// TwinCAT 3 PLC project MBIDivB_Tests
// ProgramVersion: 3.1.4024.0
// libraries:
//   MBIDivB, * (MBI Div-B)
//   Tc2_Standard, * (Beckhoff Automation GmbH)
//   Tc2_System, * (Beckhoff Automation GmbH)
//   Tc3_Module, * (Beckhoff Automation GmbH)
//   TcUnit, * (www.tcunit.org)
// project tree:
//   Example/ PRG_EXAMPLE.TcPOU
//   POUs/ FB_PlcShutdownTestable.TcPOU, PRG_TEST.TcPOU
//   / PlcTask.TcTTO
//   Tests/ FB_AnalogInputTest.TcPOU, FB_AnalogOutputTest.TcPOU, FB_CounterTimerTest.TcPOU, FB_EndPositionSwitchesTest.TcPOU, FB_FemtoAmplifierTest.TcPOU, FB_FlowMeterTest.TcPOU, FB_LedControlTest.TcPOU, FB_MultiTriggerTest.TcPOU, FB_ParameterTest.TcPOU, FB_PlcShutdownTest.TcPOU, FB_ShutterControlTest.TcPOU, FB_TimeTest.TcPOU
// (motion and I/O tree: see PLC project mbidivb)
// real-time tasks:
//   TASK PlcTask: cycle T#10ms, priority 20, ADS port 350
//   TASK PlcTask1: cycle T#1ms, priority 21, ADS port 351
// variable links:
//   MBIDivB_Tests/MBIDivB_Tests Instance <-> Device 1 (EtherCAT)/Term 1 (EK1100)/EL3102 (EL3102)
//     PlcTask Inputs/PRG_EXAMPLE.Ai1.Raw <-> AI Standard Channel 1/Value
//   MBIDivB_Tests/MBIDivB_Tests Instance <-> Device 1 (EtherCAT)/Term 1 (EK1100)/ELM3142 (ELM3142-0000)
//     PlcTask Inputs/PRG_EXAMPLE.Ai2.Raw <-> PAI Samples 1 Channel 1/Samples[0]
//   MBIDivB_Tests/MBIDivB_Tests Instance <-> Device 1 (EtherCAT)/Term 1 (EK1100)/Term 4 (EL2595)
//     PlcTask Inputs/PRG_EXAMPLE.Led1.InfoData1 <-> DOX Synchron info data/Info data 1
//     PlcTask Inputs/PRG_EXAMPLE.Led1.InfoData2 <-> DOX Synchron info data/Info data 2
//     PlcTask Inputs/PRG_EXAMPLE.Led1.StatusWord <-> DOX Status/Status
//     PlcTask Outputs/PRG_EXAMPLE.Led1.ControlWord <-> DOX Control/Control
//   MBIDivB_Tests/MBIDivB_Tests Instance <-> Device 1 (EtherCAT)/Term 1 (EK1100)/Term 5 (EL2124)
//     PlcTask Outputs/PRG_EXAMPLE.Femto1.GainBit0 <-> Channel 1/Output
//     PlcTask Outputs/PRG_EXAMPLE.Femto1.GainBit1 <-> Channel 2/Output
//     PlcTask Outputs/PRG_EXAMPLE.Femto1.GainBit2 <-> Channel 3/Output
//     PlcTask Outputs/PRG_EXAMPLE.Femto1.LowNoise <-> Channel 4/Output
//   MBIDivB_Tests/MBIDivB_Tests Instance <-> Device 1 (EtherCAT)/Term 1 (EK1100)/Term 6 (EL2124)
//     PlcTask Outputs/PRG_EXAMPLE.Femto1.DcCoupling <-> Channel 1/Output
//   MBIDivB_Tests/MBIDivB_Tests Instance <-> Device 1 (EtherCAT)/Term 1 (EK1100)/Term 7 (EL1124)
//     PlcTask Inputs/PRG_EXAMPLE.Femto1.Overload <-> Channel 1/Input

CONFIGURATION MBIDivB_Tests
    RESOURCE PLC ON TwinCAT3
        TASK PlcTask(INTERVAL := T#1ms, PRIORITY := 21);
        PROGRAM PRG_TEST WITH PlcTask : PRG_TEST;
        PROGRAM PRG_EXAMPLE WITH PlcTask : PRG_EXAMPLE;
    END_RESOURCE
END_CONFIGURATION

// ---- POUs/PRG_TEST.TcPOU

(*
    Runs all MBIDivB test suites with TcUnit. Call it from the test task
    (1 ms cycle time).
*)
PROGRAM PRG_TEST
VAR
    TimeTest : FB_TimeTest;
    ParameterTest : FB_ParameterTest;
    AnalogInputTest : FB_AnalogInputTest;
    CounterTimerTest : FB_CounterTimerTest;
    AnalogOutputTest : FB_AnalogOutputTest;
    MultiTriggerTest : FB_MultiTriggerTest;
    FlowMeterTest : FB_FlowMeterTest;
    ShutterControlTest : FB_ShutterControlTest;
    LedControlTest : FB_LedControlTest;
    FemtoAmplifierTest : FB_FemtoAmplifierTest;
    EndPositionSwitchesTest : FB_EndPositionSwitchesTest;
    PlcShutdownTest : FB_PlcShutdownTest;
END_VAR


TcUnit.RUN();

END_PROGRAM

// ---- Tests/FB_TimeTest.TcPOU

(*
    Tests of F_MsToCyclesAt, F_CyclesToMsAt and the test task's cycle time.
*)
FUNCTION_BLOCK FB_TimeTest EXTENDS TcUnit.FB_TestSuite


TaskCycleTimeIs1ms();
Converts2_4msAt1ms();
Converts1msAt0_3ms();
Converts100msAt10ms();
NonPositiveTimeGivesZero();


METHOD PRIVATE Converts100msAt10ms

TEST('Converts100msAt10ms');

AssertEquals_UDINT(Expected := 10, Actual := MBIDivB.F_MsToCyclesAt(TimeMs := 100.0, CycleTime := 100000), Message := 'cycles');
AssertEquals_REAL(Expected := 100.0, Actual := MBIDivB.F_CyclesToMsAt(Cycles := 10, CycleTime := 100000), Delta := 1.0E-6, Message := 'effective ms');

TEST_FINISHED();
END_METHOD


METHOD PRIVATE Converts1msAt0_3ms

TEST('Converts1msAt0_3ms');

AssertEquals_UDINT(Expected := 3, Actual := MBIDivB.F_MsToCyclesAt(TimeMs := 1.0, CycleTime := 3000), Message := 'cycles');
AssertEquals_REAL(Expected := 0.9, Actual := MBIDivB.F_CyclesToMsAt(Cycles := 3, CycleTime := 3000), Delta := 1.0E-6, Message := 'effective ms');

TEST_FINISHED();
END_METHOD


METHOD PRIVATE Converts2_4msAt1ms

TEST('Converts2_4msAt1ms');

AssertEquals_UDINT(Expected := 2, Actual := MBIDivB.F_MsToCyclesAt(TimeMs := 2.4, CycleTime := 10000), Message := 'cycles');
AssertEquals_REAL(Expected := 2.0, Actual := MBIDivB.F_CyclesToMsAt(Cycles := 2, CycleTime := 10000), Delta := 1.0E-6, Message := 'effective ms');

TEST_FINISHED();
END_METHOD


METHOD PRIVATE NonPositiveTimeGivesZero

TEST('NonPositiveTimeGivesZero');

AssertEquals_UDINT(Expected := 0, Actual := MBIDivB.F_MsToCyclesAt(TimeMs := 0.0, CycleTime := 10000), Message := 'zero');
AssertEquals_UDINT(Expected := 0, Actual := MBIDivB.F_MsToCyclesAt(TimeMs := -5.0, CycleTime := 10000), Message := 'negative');
AssertEquals_UDINT(Expected := 0, Actual := MBIDivB.F_MsToCyclesAt(TimeMs := 5.0, CycleTime := 0), Message := 'cycle time 0');

TEST_FINISHED();
END_METHOD


METHOD PRIVATE TaskCycleTimeIs1ms

TEST('TaskCycleTimeIs1ms');

AssertEquals_UDINT(Expected := 10000, Actual := MBIDivB.F_GetTaskCycleTime(),
    Message := 'The test task must run at 1 ms; the other suites assume it');

TEST_FINISHED();
END_METHOD

END_FUNCTION_BLOCK

// ---- Tests/FB_ParameterTest.TcPOU

(*
    Checks that the library parameter overrides of this test project take
    effect (task 10.1). Expected overrides in the Library Manager:
    CT_CHANNELS 4, CT_BUFFER_LENGTH 1000, AO_WAVEFORM_LENGTH 1000,
    FLOW_BUFFER_LENGTH 100.
*)
FUNCTION_BLOCK FB_ParameterTest EXTENDS TcUnit.FB_TestSuite
VAR
    Ct : MBIDivB.FB_CounterTimer;
    Ao : MBIDivB.FB_AnalogOutput;
END_VAR


OverridesSetArrayBounds();


METHOD PRIVATE OverridesSetArrayBounds

TEST('OverridesSetArrayBounds');

// Element counts from the array sizes (UPPER_BOUND only works on
// variable-length arrays in TwinCAT 3.1.4024).
AssertEquals_UDINT(Expected := 4, Actual := TO_UDINT(SIZEOF(Ct.Channel) / SIZEOF(Ct.Channel[1])), Message := 'CT_CHANNELS');
AssertEquals_UDINT(Expected := 1000, Actual := TO_UDINT(SIZEOF(Ct.Channel[1].Data) / SIZEOF(Ct.Channel[1].Data[1])), Message := 'CT_BUFFER_LENGTH');
AssertEquals_UDINT(Expected := 1000, Actual := TO_UDINT(SIZEOF(Ao.Data) / SIZEOF(Ao.Data[1])), Message := 'AO_WAVEFORM_LENGTH');
AssertEquals_UDINT(Expected := 100, Actual := MBIDivB.GVL_Param.FLOW_BUFFER_LENGTH, Message := 'FLOW_BUFFER_LENGTH');

TEST_FINISHED();
END_METHOD

END_FUNCTION_BLOCK

// ---- Tests/FB_AnalogInputTest.TcPOU

(*
    Tests of FB_AnalogInput16/32 (specs/analog-input).
*)
FUNCTION_BLOCK FB_AnalogInputTest EXTENDS TcUnit.FB_TestSuite
VAR
    AiNegative : MBIDivB.FB_AnalogInput16;
    AiElmNominal : MBIDivB.FB_AnalogInput32;
    AiElmPreset : MBIDivB.FB_AnalogInput32;
    AiZeroScale : MBIDivB.FB_AnalogInput16;
    AiConstant : MBIDivB.FB_AnalogInput16;
    AiReduced : MBIDivB.FB_AnalogInput16;
    AiSizeZero : MBIDivB.FB_AnalogInput16;
    AiOverrange : MBIDivB.FB_AnalogInput16;
    AiUnlinked : MBIDivB.FB_AnalogInput32;
    AiRestartStep : MBIDivB.FB_AnalogInput16;
    AiRestartSettings : MBIDivB.FB_AnalogInput32;
END_VAR


NegativeValue16Bit();
ElmNominalFullScale();
ElmExtendedPreset();
ZeroRawFullScaleRejected();
ConstantInputFiltered();
FilterSizeReducedRestarts();
FilterSizeZeroClampedToOne();
OverrangeSetAndCleared();
UnlinkedStatusBitsNoError();
RestartAfterStep();
RestartKeepsSettings();


METHOD PRIVATE ConstantInputFiltered
VAR
    Cycle : INT;
END_VAR

TEST('ConstantInputFiltered');

AiConstant.SetScale(RawFullScale := 1, ValueFullScale := 1.0);
AiConstant.Cfg.FilterSize := 10;
AiConstant.Raw := 2;
FOR Cycle := 1 TO 25 DO
    AiConstant();
END_FOR
AssertEquals_REAL(Expected := 2.0, Actual := AiConstant.Status.ValueFiltered, Delta := 1.0E-6, Message := 'ValueFiltered');

TEST_FINISHED();
END_METHOD


METHOD PRIVATE ElmExtendedPreset

TEST('ElmExtendedPreset');

AiElmPreset.SetScalePreset(Preset := MBIDivB.E_AiScalePreset.ELM3XXX_EXTENDED, NominalFullScale := 10.0);
AiElmPreset.Raw := 7812500;
AiElmPreset();
AssertEquals_REAL(Expected := 10.0, Actual := AiElmPreset.Status.Value, Delta := 1.0E-5, Message := 'nominal');
AiElmPreset.Raw := 8388607;
AiElmPreset();
AssertEquals_REAL(Expected := 10.737, Actual := AiElmPreset.Status.Value, Delta := 0.001, Message := 'technical full scale');

TEST_FINISHED();
END_METHOD


METHOD PRIVATE ElmNominalFullScale

TEST('ElmNominalFullScale');

AiElmNominal.SetScale(RawFullScale := 7812500, ValueFullScale := 10.0);
AiElmNominal.Raw := 7812500;
AiElmNominal();
AssertEquals_REAL(Expected := 10.0, Actual := AiElmNominal.Status.Value, Delta := 1.0E-5, Message := 'Value');
AssertEquals_DINT(Expected := 7812500, Actual := AiElmNominal.Status.RawFullScale, Message := 'RawFullScale');
AssertEquals_REAL(Expected := 10.0, Actual := AiElmNominal.Status.ValueFullScale, Delta := 1.0E-6, Message := 'ValueFullScale');

TEST_FINISHED();
END_METHOD


METHOD PRIVATE FilterSizeReducedRestarts
VAR
    Cycle : INT;
END_VAR

TEST('FilterSizeReducedRestarts');

AiReduced.SetScale(RawFullScale := 1, ValueFullScale := 1.0);
AiReduced.Cfg.FilterSize := 1000;
AiReduced.Raw := 3;
FOR Cycle := 1 TO 100 DO
    AiReduced();
END_FOR
AiReduced.Cfg.FilterSize := 10;
AiReduced.Raw := 1;
AiReduced();
AssertEquals_REAL(Expected := 1.0, Actual := AiReduced.Status.ValueFiltered, Delta := 1.0E-6, Message := 'no contribution from older samples');

TEST_FINISHED();
END_METHOD


METHOD PRIVATE FilterSizeZeroClampedToOne

TEST('FilterSizeZeroClampedToOne');

AiSizeZero.SetScale(RawFullScale := 1, ValueFullScale := 1.0);
AiSizeZero.Cfg.FilterSize := 0;
AiSizeZero.Raw := 4;
AiSizeZero();
AssertEquals_DINT(Expected := 1, Actual := AiSizeZero.Cfg.FilterSize, Message := 'FilterSize written back');
AssertEquals_REAL(Expected := 4.0, Actual := AiSizeZero.Status.ValueFiltered, Delta := 1.0E-6, Message := 'ValueFiltered');

TEST_FINISHED();
END_METHOD


METHOD PRIVATE NegativeValue16Bit

TEST('NegativeValue16Bit');

AiNegative.SetScalePreset(Preset := MBIDivB.E_AiScalePreset.EL31XX_LEGACY, NominalFullScale := 10.0);
AiNegative.Raw := -16384;
AiNegative();
AssertEquals_REAL(Expected := -5.0, Actual := AiNegative.Status.Value, Delta := 0.001, Message := 'Value');
AssertEquals_DINT(Expected := -16384, Actual := AiNegative.Status.Raw, Message := 'Raw');

TEST_FINISHED();
END_METHOD


METHOD PRIVATE OverrangeSetAndCleared

TEST('OverrangeSetAndCleared');

AiOverrange.Overrange := TRUE;
AiOverrange();
AssertTrue(Condition := AiOverrange.Status.Error, Message := 'Error while set');
AssertTrue(Condition := FIND(AiOverrange.Status.ErrorText, 'overrange') > 0, Message := 'ErrorText mentions overrange');
AiOverrange.Overrange := FALSE;
AiOverrange();
AssertFalse(Condition := AiOverrange.Status.Error, Message := 'Error cleared');
AssertEquals_STRING(Expected := '', Actual := AiOverrange.Status.ErrorText, Message := 'ErrorText cleared');

TEST_FINISHED();
END_METHOD


METHOD PRIVATE RestartAfterStep
VAR
    Cycle : INT;
    Wrong : INT;
END_VAR

TEST('RestartAfterStep');

AiRestartStep.SetScale(RawFullScale := 1000, ValueFullScale := 1.0);
AiRestartStep.Cfg.FilterSize := 10;
AiRestartStep.Raw := 1000;
FOR Cycle := 1 TO 15 DO
    AiRestartStep();
END_FOR
AiRestartStep.RestartFilter();
AiRestartStep.Raw := 3000;
FOR Cycle := 1 TO 12 DO
    AiRestartStep();
    IF ABS(AiRestartStep.Status.ValueFiltered - 3.0) > 1.0E-6 THEN
        Wrong := Wrong + 1;
    END_IF
END_FOR
AssertEquals_INT(Expected := 0, Actual := Wrong, Message := 'calls with ValueFiltered <> 3.0 V after the restart');

TEST_FINISHED();
END_METHOD


METHOD PRIVATE RestartKeepsSettings

TEST('RestartKeepsSettings');

AiRestartSettings.SetScale(RawFullScale := 7812500, ValueFullScale := 10.0);
AiRestartSettings.Cfg.FilterSize := 20;
AiRestartSettings.Raw := 3906250;
AiRestartSettings();
AiRestartSettings.RestartFilter();
AiRestartSettings();
AssertEquals_DINT(Expected := 20, Actual := AiRestartSettings.Cfg.FilterSize, Message := 'FilterSize');
AssertEquals_DINT(Expected := 7812500, Actual := AiRestartSettings.Status.RawFullScale, Message := 'RawFullScale');
AssertEquals_REAL(Expected := 10.0, Actual := AiRestartSettings.Status.ValueFullScale, Delta := 1.0E-6, Message := 'ValueFullScale');
AssertEquals_REAL(Expected := 5.0, Actual := AiRestartSettings.Status.Value, Delta := 1.0E-5, Message := 'Value');

TEST_FINISHED();
END_METHOD


METHOD PRIVATE UnlinkedStatusBitsNoError

TEST('UnlinkedStatusBitsNoError');

AiUnlinked.Raw := 1000;
AiUnlinked();
AssertFalse(Condition := AiUnlinked.Status.Error, Message := 'Error');

TEST_FINISHED();
END_METHOD


METHOD PRIVATE ZeroRawFullScaleRejected
VAR
    Accepted : BOOL;
END_VAR

TEST('ZeroRawFullScaleRejected');

AiZeroScale.SetScale(RawFullScale := 32767, ValueFullScale := 10.0);
Accepted := AiZeroScale.SetScale(RawFullScale := 0, ValueFullScale := 5.0);
AiZeroScale.Raw := 16384;
AiZeroScale();
AssertFalse(Condition := Accepted, Message := 'SetScale must return FALSE');
AssertTrue(Condition := AiZeroScale.Status.Error, Message := 'Error');
AssertTrue(Condition := FIND(AiZeroScale.Status.ErrorText, 'RawFullScale') > 0, Message := 'ErrorText names RawFullScale');
AssertEquals_REAL(Expected := 5.0, Actual := AiZeroScale.Status.Value, Delta := 0.001, Message := 'previous scaling kept');

TEST_FINISHED();
END_METHOD

END_FUNCTION_BLOCK

// ---- Tests/FB_CounterTimerTest.TcPOU

(*
    Tests of FB_CounterTimer (specs/counter-timer) and of the command
    handshake and error rules (specs/ads-interface) on this block.
    Needs CT_CHANNELS >= 4.
*)
FUNCTION_BLOCK FB_CounterTimerTest EXTENDS TcUnit.FB_TestSuite
VAR
    CtSync : MBIDivB.FB_CounterTimer;
    CtTooMany : MBIDivB.FB_CounterTimer;
    CtLinear : MBIDivB.FB_CounterTimer;
    CtLatency : MBIDivB.FB_CounterTimer;
    CtTrigger : MBIDivB.FB_CounterTimer;
    CtMissed : MBIDivB.FB_CounterTimer;
    CtProgress : MBIDivB.FB_CounterTimer;
    CtStop : MBIDivB.FB_CounterTimer;
    CtRunning : MBIDivB.FB_CounterTimer;
    CtHandshake : MBIDivB.FB_CounterTimer;
    CtErrorClear : MBIDivB.FB_CounterTimer;
    CtCfgChange : MBIDivB.FB_CounterTimer;
END_VAR


SynchronousPoints();
TooManyPointsRejected();
LinearInputMean();
WindowsWithLatency();
ThreeTriggerPoints();
EverySecondEdgeMissed();
ProgressDuringAcquisition();
StopKeepsPoints();
StartWhileRunningRejected();
StartHandshake();
ErrorClearedByAcceptedStart();
ConfigChangeDuringRun();


METHOD PRIVATE ConfigChangeDuringRun
VAR
    Cycle : INT;
END_VAR

TEST('ConfigChangeDuringRun');

CtCfgChange.Cfg.IntegrationTimeMs := 2.0;
CtCfgChange.Cfg.Points := 2;
CtCfgChange.Cmd.Start := TRUE;
CtCfgChange();
CtCfgChange.Cfg.IntegrationTimeMs := 100.0;
FOR Cycle := 1 TO 4 DO
    CtCfgChange();
END_FOR
AssertEquals_DINT(Expected := 2, Actual := CtCfgChange.Status.PointsDone, Message := 'started integration time kept');
AssertEquals_REAL(Expected := 2.0, Actual := CtCfgChange.Status.IntegrationTimeMs, Delta := 1.0E-6, Message := 'effective time');

TEST_FINISHED();
END_METHOD


METHOD PRIVATE ErrorClearedByAcceptedStart

TEST('ErrorClearedByAcceptedStart');

CtErrorClear.Cfg.IntegrationTimeMs := 0.0;
CtErrorClear.Cmd.Start := TRUE;
CtErrorClear();
AssertFalse(Condition := CtErrorClear.Cmd.Start, Message := 'flag cleared');
AssertEquals_INT(Expected := 0, Actual := CtErrorClear.Status.State, Message := 'stays idle');
AssertTrue(Condition := CtErrorClear.Status.Error, Message := 'Error');
AssertTrue(Condition := FIND(CtErrorClear.Status.ErrorText, 'IntegrationTimeMs') > 0, Message := 'names IntegrationTimeMs');
CtErrorClear.Cfg.IntegrationTimeMs := 10.0;
CtErrorClear.Cmd.Start := TRUE;
CtErrorClear();
AssertFalse(Condition := CtErrorClear.Status.Error, Message := 'Error cleared');
AssertEquals_STRING(Expected := '', Actual := CtErrorClear.Status.ErrorText, Message := 'ErrorText cleared');

TEST_FINISHED();
END_METHOD


METHOD PRIVATE EverySecondEdgeMissed
VAR
    Cycle : INT;
END_VAR

TEST('EverySecondEdgeMissed');

CtMissed.Cfg.StartMode := 1;
CtMissed.Cfg.IntegrationTimeMs := 8.0;
CtMissed.Cfg.Points := 100;
CtMissed.Start();
FOR Cycle := 0 TO 50 DO
    CtMissed(Gate := Cycle > 0 AND Cycle MOD 5 = 0);
END_FOR
// Edges at 5, 15, 25, 35, 45 start windows; 10, 20, 30, 40, 50 are missed.
AssertEquals_UDINT(Expected := 5, Actual := CtMissed.Status.MissedTriggers, Message := 'MissedTriggers');
AssertEquals_DINT(Expected := 4, Actual := CtMissed.Status.PointsDone, Message := 'PointsDone');

TEST_FINISHED();
END_METHOD


METHOD PRIVATE LinearInputMean
VAR
    Cycle : INT;
END_VAR

TEST('LinearInputMean');

CtLinear.Cfg.IntegrationTimeMs := 4.0;
CtLinear.Cfg.Points := 1;
CtLinear.Cmd.Start := TRUE;
CtLinear();   // start cycle, window 1 starts in the next cycle
FOR Cycle := 1 TO 4 DO
    CtLinear.Channel[1].Input := INT_TO_REAL(Cycle);
    CtLinear();
END_FOR
AssertEquals_REAL(Expected := 2.5, Actual := CtLinear.Channel[1].Data[1], Delta := 1.0E-6, Message := 'mean of 1..4');
AssertEquals_INT(Expected := 0, Actual := CtLinear.Status.State, Message := 'idle after the last point');

TEST_FINISHED();
END_METHOD


METHOD PRIVATE ProgressDuringAcquisition
VAR
    Cycle : INT;
END_VAR

TEST('ProgressDuringAcquisition');

CtProgress.Cfg.IntegrationTimeMs := 1.0;
CtProgress.Cfg.Points := 10;
CtProgress.Cmd.Start := TRUE;
FOR Cycle := 0 TO 4 DO
    CtProgress();
END_FOR
AssertEquals_DINT(Expected := 4, Actual := CtProgress.Status.PointsDone, Message := 'PointsDone');
AssertTrue(Condition := CtProgress.Status.State <> 0, Message := 'not idle');

TEST_FINISHED();
END_METHOD


METHOD PRIVATE StartHandshake
VAR
    ReadBeforeCycle : BOOL;
END_VAR

TEST('StartHandshake');

CtHandshake.Cmd.Start := TRUE;
ReadBeforeCycle := CtHandshake.Cmd.Start;
CtHandshake();
AssertTrue(Condition := ReadBeforeCycle, Message := 'flag reads TRUE before the PLC cycle');
AssertFalse(Condition := CtHandshake.Cmd.Start, Message := 'flag cleared');
AssertEquals_INT(Expected := 1, Actual := CtHandshake.Status.State, Message := 'running state when the flag reads FALSE');
AssertEquals_STRING(Expected := 'INTEGRATING', Actual := CtHandshake.Status.StateText, Message := 'TO_STRING of E_CtState');

TEST_FINISHED();
END_METHOD


METHOD PRIVATE StartWhileRunningRejected
VAR
    Cycle : INT;
END_VAR

TEST('StartWhileRunningRejected');

CtRunning.Cfg.IntegrationTimeMs := 5.0;
CtRunning.Cfg.Points := 2;
CtRunning.Cmd.Start := TRUE;
CtRunning();
CtRunning();
CtRunning.Cmd.Start := TRUE;
CtRunning();
AssertFalse(Condition := CtRunning.Cmd.Start, Message := 'flag cleared');
AssertTrue(Condition := CtRunning.Status.Error, Message := 'Error');
AssertEquals_INT(Expected := 1, Actual := CtRunning.Status.State, Message := 'still integrating');
FOR Cycle := 1 TO 20 DO
    CtRunning();
END_FOR
AssertEquals_DINT(Expected := 2, Actual := CtRunning.Status.PointsDone, Message := 'running acquisition completed');

TEST_FINISHED();
END_METHOD


METHOD PRIVATE StopKeepsPoints
VAR
    Cycle : INT;
    Point : INT;
    Before : ARRAY[1..5] OF REAL;
END_VAR

TEST('StopKeepsPoints');

CtStop.Cfg.IntegrationTimeMs := 2.0;
CtStop.Cfg.Points := 10;
CtStop.Cmd.Start := TRUE;
FOR Cycle := 0 TO 11 DO   // points 1-5 in cycles 1-10, cycle 11 starts point 6
    CtStop.Channel[1].Input := INT_TO_REAL(Cycle);
    CtStop();
END_FOR
FOR Point := 1 TO 5 DO
    Before[Point] := CtStop.Channel[1].Data[Point];
END_FOR
CtStop.Cmd.Stop := TRUE;
CtStop();
AssertEquals_INT(Expected := 0, Actual := CtStop.Status.State, Message := 'idle');
AssertEquals_DINT(Expected := 5, Actual := CtStop.Status.PointsDone, Message := 'PointsDone');
FOR Point := 1 TO 5 DO
    AssertEquals_REAL(Expected := Before[Point], Actual := CtStop.Channel[1].Data[Point], Delta := 0.0, Message := 'point unchanged');
END_FOR

TEST_FINISHED();
END_METHOD


METHOD PRIVATE SynchronousPoints
VAR
    Cycle : INT;
    Channel : INT;
    Point : INT;
END_VAR

TEST('SynchronousPoints');

CtSync.Cfg.IntegrationTimeMs := 2.0;
CtSync.Cfg.Points := 10;
CtSync.Start();
FOR Cycle := 0 TO 30 DO
    FOR Channel := 1 TO 4 DO
        CtSync.Channel[Channel].Input := INT_TO_REAL(Channel * 1000 + Cycle);
    END_FOR
    CtSync();
END_FOR
AssertEquals_DINT(Expected := 10, Actual := CtSync.Status.PointsDone, Message := 'PointsDone');
FOR Point := 1 TO 10 DO
    FOR Channel := 2 TO 4 DO
        // Same cycles: the channel offset is the only difference.
        AssertEquals_REAL(Expected := CtSync.Channel[1].Data[Point] + INT_TO_REAL((Channel - 1) * 1000),
            Actual := CtSync.Channel[Channel].Data[Point], Delta := 0.01, Message := 'point from the same cycles');
    END_FOR
END_FOR

TEST_FINISHED();
END_METHOD


METHOD PRIVATE ThreeTriggerPoints
VAR
    Cycle : INT;
END_VAR

TEST('ThreeTriggerPoints');

CtTrigger.Cfg.StartMode := 1;
CtTrigger.Cfg.IntegrationTimeMs := 3.0;
CtTrigger.Cfg.Points := 3;
CtTrigger.Start();
AssertEquals_INT(Expected := 3, Actual := CtTrigger.Status.State, Message := 'WAIT_TRIGGER after start');
FOR Cycle := 0 TO 30 DO
    CtTrigger.Channel[1].Input := INT_TO_REAL(Cycle);
    CtTrigger(Gate := Cycle = 5 OR Cycle = 15 OR Cycle = 25);
END_FOR
AssertEquals_DINT(Expected := 3, Actual := CtTrigger.Status.PointsDone, Message := 'PointsDone');
AssertEquals_REAL(Expected := 6.0, Actual := CtTrigger.Channel[1].Data[1], Delta := 1.0E-6, Message := 'point 1 from the edge cycle on');
AssertEquals_REAL(Expected := 16.0, Actual := CtTrigger.Channel[1].Data[2], Delta := 1.0E-6, Message := 'point 2');
AssertEquals_REAL(Expected := 26.0, Actual := CtTrigger.Channel[1].Data[3], Delta := 1.0E-6, Message := 'point 3');
AssertEquals_UDINT(Expected := 0, Actual := CtTrigger.Status.MissedTriggers, Message := 'MissedTriggers');
AssertEquals_INT(Expected := 0, Actual := CtTrigger.Status.State, Message := 'idle');

TEST_FINISHED();
END_METHOD


METHOD PRIVATE TooManyPointsRejected

TEST('TooManyPointsRejected');

CtTooMany.Cfg.Points := UDINT_TO_DINT(MBIDivB.GVL_Param.CT_BUFFER_LENGTH) + 1;
CtTooMany.Cmd.Start := TRUE;
CtTooMany();
AssertFalse(Condition := CtTooMany.Cmd.Start, Message := 'flag cleared');
AssertEquals_INT(Expected := 0, Actual := CtTooMany.Status.State, Message := 'stays idle');
AssertTrue(Condition := CtTooMany.Status.Error, Message := 'Error');
AssertTrue(Condition := FIND(CtTooMany.Status.ErrorText, 'Points') > 0, Message := 'names Points');
AssertTrue(Condition := FIND(CtTooMany.Status.ErrorText, UDINT_TO_STRING(MBIDivB.GVL_Param.CT_BUFFER_LENGTH)) > 0, Message := 'names the buffer length');

TEST_FINISHED();
END_METHOD


METHOD PRIVATE WindowsWithLatency
VAR
    Cycle : INT;
    IdleAfter18 : BOOL;
END_VAR

TEST('WindowsWithLatency');

CtLatency.Cfg.IntegrationTimeMs := 5.0;
CtLatency.Cfg.LatencyTimeMs := 2.0;
CtLatency.Cfg.Points := 3;
CtLatency.Cmd.Start := TRUE;
FOR Cycle := 0 TO 19 DO
    CtLatency.Channel[1].Input := INT_TO_REAL(Cycle);
    CtLatency();
    IF Cycle = 18 THEN
        IdleAfter18 := CtLatency.Status.State = 0;
    END_IF
END_FOR
AssertEquals_REAL(Expected := 3.0, Actual := CtLatency.Channel[1].Data[1], Delta := 1.0E-6, Message := 'window 1 = cycles 1-5');
AssertEquals_REAL(Expected := 10.0, Actual := CtLatency.Channel[1].Data[2], Delta := 1.0E-6, Message := 'window 2 = cycles 8-12');
AssertEquals_REAL(Expected := 17.0, Actual := CtLatency.Channel[1].Data[3], Delta := 1.0E-6, Message := 'window 3 = cycles 15-19');
AssertFalse(Condition := IdleAfter18, Message := 'running until cycle 19');
AssertEquals_INT(Expected := 0, Actual := CtLatency.Status.State, Message := 'idle after the third window');
AssertEquals_REAL(Expected := 5.0, Actual := CtLatency.Status.IntegrationTimeMs, Delta := 1.0E-6, Message := 'effective integration time');
AssertEquals_REAL(Expected := 2.0, Actual := CtLatency.Status.LatencyTimeMs, Delta := 1.0E-6, Message := 'effective latency time');

TEST_FINISHED();
END_METHOD

END_FUNCTION_BLOCK

// ---- Tests/FB_AnalogOutputTest.TcPOU

(*
    Tests of FB_AnalogOutput (specs/analog-output). Needs AO_WAVEFORM_LENGTH >= 4.
*)
FUNCTION_BLOCK FB_AnalogOutputTest EXTENDS TcUnit.FB_TestSuite
VAR
    AoBack : MBIDivB.FB_AnalogOutput;
    AoDuration : MBIDivB.FB_AnalogOutput;
    AoReversal : MBIDivB.FB_AnalogOutput;
    AoReached : MBIDivB.FB_AnalogOutput;
    AoZeroVelocity : MBIDivB.FB_AnalogOutput;
    AoLimit : MBIDivB.FB_AnalogOutput;
    AoFull : MBIDivB.FB_AnalogOutput;
    AoStep : MBIDivB.FB_AnalogOutput;
    AoEndless : MBIDivB.FB_AnalogOutput;
    AoRampStart : MBIDivB.FB_AnalogOutput;
    AoBoot : MBIDivB.FB_AnalogOutput;
    AoProgress : MBIDivB.FB_AnalogOutput;
    AoX : MBIDivB.FB_AnalogOutput;
    AoY : MBIDivB.FB_AnalogOutput;
    AoRecord : MBIDivB.FB_AnalogOutput;
    CtRecord : MBIDivB.FB_CounterTimer;
END_VAR


BackToRampMode();
RampDuration();
SetpointChangedMidRamp();
SetpointReachedFlag();
ZeroVelocityKeepsPrevious();
SetpointAboveLimit();
FullPositiveOutput();
StepTime4x10Cycles();
EndlessRepetition();
StartInRampModeRejected();
IdleAtStartInWaveformMode();
WaveformProgress();
TwoOutputsInLockstep();
PresentValueRecorded();


METHOD PRIVATE BackToRampMode
VAR
    Cycle : INT;
END_VAR

TEST('BackToRampMode');

AoBack.Cfg.Mode := 1;
AoBack.Data[1] := 3.0;
AoBack.Cfg.WaveformPoints := 1;
AoBack.Cfg.Repeats := 0;
AoBack.Cmd.Start := TRUE;
FOR Cycle := 1 TO 5 DO
    AoBack();
END_FOR
AssertEquals_REAL(Expected := 3.0, Actual := AoBack.Status.Value, Delta := 1.0E-6, Message := 'waveform output');
AoBack.Cfg.Setpoint := 0.0;
AoBack.Cfg.VelocityVPerS := 1.0;
AoBack.Cfg.Mode := 0;
AoBack();
AssertEquals_INT(Expected := 0, Actual := AoBack.Status.State, Message := 'ramp state, waveform stopped');
AssertEquals_REAL(Expected := 2.999, Actual := AoBack.Status.Value, Delta := 1.0E-5, Message := 'ramps from 3.0 V');
FOR Cycle := 1 TO 3000 DO
    AoBack();
END_FOR
AssertEquals_REAL(Expected := 0.0, Actual := AoBack.Status.Value, Delta := 0.0, Message := 'at setpoint');

TEST_FINISHED();
END_METHOD


METHOD PRIVATE EndlessRepetition
VAR
    Cycle : INT;
END_VAR

TEST('EndlessRepetition');

AoEndless.Cfg.Mode := 1;
AoEndless.Data[1] := 1.0;
AoEndless.Data[2] := -1.0;
AoEndless.Cfg.WaveformPoints := 2;
AoEndless.Cfg.Repeats := 0;
AoEndless.Cmd.Start := TRUE;
FOR Cycle := 1 TO 1000 DO
    AoEndless();
END_FOR
AssertEquals_INT(Expected := 2, Actual := AoEndless.Status.State, Message := 'still playing');
AssertEquals_DINT(Expected := 500, Actual := AoEndless.Status.RepeatsDone, Message := 'RepeatsDone');
AoEndless.Cmd.Stop := TRUE;
AoEndless();
AssertEquals_INT(Expected := 1, Actual := AoEndless.Status.State, Message := 'stopped');

TEST_FINISHED();
END_METHOD


METHOD PRIVATE FullPositiveOutput
VAR
    Cycle : INT;
END_VAR

TEST('FullPositiveOutput');

AoFull.Cfg.VelocityVPerS := 1000.0;
AoFull.Cfg.Setpoint := 10.0;
FOR Cycle := 1 TO 20 DO
    AoFull();
END_FOR
AssertEquals_INT(Expected := 32767, Actual := AoFull.Raw, Message := 'Raw output');
AssertEquals_INT(Expected := 32767, Actual := AoFull.Status.Raw, Message := 'Status.Raw');

TEST_FINISHED();
END_METHOD


METHOD PRIVATE IdleAtStartInWaveformMode
VAR
    Cycle : INT;
END_VAR

TEST('IdleAtStartInWaveformMode');

AoBoot.Cfg.Mode := 1;
AoBoot.Data[1] := 7.0;
FOR Cycle := 1 TO 10 DO
    AoBoot();
END_FOR
AssertEquals_INT(Expected := 1, Actual := AoBoot.Status.State, Message := 'WAVEFORM_IDLE');
AssertEquals_REAL(Expected := 0.0, Actual := AoBoot.Status.Value, Delta := 0.0, Message := 'holds the initial value');

TEST_FINISHED();
END_METHOD


METHOD PRIVATE PresentValueRecorded
VAR
    Cycle : INT;
END_VAR

TEST('PresentValueRecorded');

AoRecord.Cfg.VelocityVPerS := 1000.0;
AoRecord.Cfg.Setpoint := 1.25;
FOR Cycle := 1 TO 5 DO
    AoRecord();
END_FOR
CtRecord.Cfg.IntegrationTimeMs := 1.0;
CtRecord.Cfg.Points := 1;
CtRecord.Start();
FOR Cycle := 1 TO 2 DO
    AoRecord();
    CtRecord.Channel[1].Input := AoRecord.Status.Value;
    CtRecord();
END_FOR
AssertEquals_REAL(Expected := 1.25, Actual := CtRecord.Channel[1].Data[1], Delta := 0.0, Message := 'acquires the output value');
AssertEquals_INT(Expected := 4096, Actual := AoRecord.Status.Raw, Message := 'Raw = 1.25 V x 32767 / 10 V');

TEST_FINISHED();
END_METHOD


METHOD PRIVATE RampDuration
VAR
    Cycle : INT;
    MaxValue : REAL;
    ReachedAt : INT;
END_VAR

TEST('RampDuration');

AoDuration.Cfg.VelocityVPerS := 2.0;
AoDuration.Cfg.Setpoint := 1.0;
ReachedAt := -1;
FOR Cycle := 1 TO 600 DO
    AoDuration();
    MaxValue := MAX(MaxValue, AoDuration.Status.Value);
    IF ReachedAt < 0 AND AoDuration.Status.Value = 1.0 THEN
        ReachedAt := Cycle;
    END_IF
END_FOR
AssertEquals_INT(Expected := 500, Actual := ReachedAt, Message := 'reached after 0.5 s');
AssertEquals_REAL(Expected := 1.0, Actual := MaxValue, Delta := 0.0, Message := 'no overshoot');

TEST_FINISHED();
END_METHOD


METHOD PRIVATE SetpointAboveLimit
VAR
    Cycle : INT;
END_VAR

TEST('SetpointAboveLimit');

AoLimit.Cfg.LimitMax := 5.0;
AoLimit.Cfg.VelocityVPerS := 100.0;
AoLimit.Cfg.Setpoint := 8.0;
FOR Cycle := 1 TO 100 DO
    AoLimit();
END_FOR
AssertEquals_REAL(Expected := 5.0, Actual := AoLimit.Status.Value, Delta := 0.0, Message := 'output at the limit');
AssertEquals_REAL(Expected := 8.0, Actual := AoLimit.Cfg.Setpoint, Delta := 0.0, Message := 'Cfg.Setpoint keeps the written value');
AssertTrue(Condition := AoLimit.Status.Limited, Message := 'Limited');

TEST_FINISHED();
END_METHOD


METHOD PRIVATE SetpointChangedMidRamp
VAR
    Cycle : INT;
    Previous : REAL;
    MaxStep : REAL;
END_VAR

TEST('SetpointChangedMidRamp');

AoReversal.Cfg.VelocityVPerS := 1.0;
AoReversal.Cfg.Setpoint := 2.0;
FOR Cycle := 1 TO 1500 DO
    AoReversal();
END_FOR
AssertEquals_REAL(Expected := 1.5, Actual := AoReversal.Status.Value, Delta := 1.0E-4, Message := 'ramping at 1.5 V');
Previous := AoReversal.Status.Value;
AoReversal.Cfg.Setpoint := 0.0;
FOR Cycle := 1 TO 2000 DO
    AoReversal();
    MaxStep := MAX(MaxStep, ABS(AoReversal.Status.Value - Previous));
    Previous := AoReversal.Status.Value;
END_FOR
AssertTrue(Condition := MaxStep <= 0.00101, Message := 'no step larger than velocity x cycle time');
AssertEquals_REAL(Expected := 0.0, Actual := AoReversal.Status.Value, Delta := 0.0, Message := 'reaches 0 V');

TEST_FINISHED();
END_METHOD


METHOD PRIVATE SetpointReachedFlag
VAR
    Cycle : INT;
END_VAR

TEST('SetpointReachedFlag');

AoReached.Cfg.VelocityVPerS := 1.0;
AoReached.Cfg.Setpoint := 0.01;
AoReached();
AssertFalse(Condition := AoReached.Status.SetpointReached, Message := 'FALSE while ramping');
FOR Cycle := 1 TO 20 DO
    AoReached();
END_FOR
AssertTrue(Condition := AoReached.Status.SetpointReached, Message := 'TRUE at the setpoint');

TEST_FINISHED();
END_METHOD


METHOD PRIVATE StartInRampModeRejected

TEST('StartInRampModeRejected');

AoRampStart.Cmd.Start := TRUE;
AoRampStart();
AssertFalse(Condition := AoRampStart.Cmd.Start, Message := 'flag cleared');
AssertTrue(Condition := AoRampStart.Status.Error, Message := 'Error');
AssertTrue(Condition := FIND(AoRampStart.Status.ErrorText, 'Mode') > 0, Message := 'names the mode');
AssertEquals_INT(Expected := 0, Actual := AoRampStart.Status.State, Message := 'state unchanged');

TEST_FINISHED();
END_METHOD


METHOD PRIVATE StepTime4x10Cycles
VAR
    Cycle : INT;
    Wrong : INT;
END_VAR

TEST('StepTime4x10Cycles');

AoStep.Cfg.Mode := 1;
AoStep.Data[1] := 1.0;
AoStep.Data[2] := 2.0;
AoStep.Data[3] := 3.0;
AoStep.Data[4] := 4.0;
AoStep.Cfg.WaveformPoints := 4;
AoStep.Cfg.StepTimeMs := 10.0;
AoStep.Cfg.Repeats := 1;
AoStep.Cmd.Start := TRUE;
FOR Cycle := 0 TO 39 DO
    AoStep();
    IF AoStep.Status.Value <> INT_TO_REAL(Cycle / 10 + 1) THEN
        Wrong := Wrong + 1;
    END_IF
END_FOR
AssertEquals_INT(Expected := 0, Actual := Wrong, Message := 'each element for 10 cycles');
AssertEquals_INT(Expected := 1, Actual := AoStep.Status.State, Message := 'idle after 40 cycles');
FOR Cycle := 1 TO 10 DO
    AoStep();
END_FOR
AssertEquals_REAL(Expected := 4.0, Actual := AoStep.Status.Value, Delta := 0.0, Message := 'holds element 4');

TEST_FINISHED();
END_METHOD


METHOD PRIVATE TwoOutputsInLockstep
VAR
    Cycle : INT;
    Point : INT;
    Mismatch : INT;
END_VAR

TEST('TwoOutputsInLockstep');

AoX.Cfg.Mode := 1;
AoY.Cfg.Mode := 1;
FOR Point := 1 TO 4 DO
    AoX.Data[Point] := INT_TO_REAL(Point);
    AoY.Data[Point] := INT_TO_REAL(-Point);
END_FOR
AoX.Cfg.WaveformPoints := 4;
AoY.Cfg.WaveformPoints := 4;
AoX.Cfg.StepTimeMs := 3.0;
AoY.Cfg.StepTimeMs := 3.0;
AoX();
AoY();
AoX.Start();
AoY.Start();
FOR Cycle := 1 TO 12 DO
    AoX();
    AoY();
    IF AoX.Status.Index <> AoY.Status.Index OR AoX.Status.Value <> -AoY.Status.Value THEN
        Mismatch := Mismatch + 1;
    END_IF
END_FOR
AssertEquals_INT(Expected := 0, Actual := Mismatch, Message := 'element k in the same cycle');

TEST_FINISHED();
END_METHOD


METHOD PRIVATE WaveformProgress
VAR
    Cycle : INT;
END_VAR

TEST('WaveformProgress');

AoProgress.Cfg.Mode := 1;
AoProgress.Cfg.WaveformPoints := 4;
AoProgress.Cfg.StepTimeMs := 1.0;
AoProgress.Cfg.Repeats := 3;
AoProgress.Cmd.Start := TRUE;
FOR Cycle := 0 TO 6 DO   // pass 1 in cycles 0-3, pass 2 element 3 in cycle 6
    AoProgress();
END_FOR
AssertEquals_DINT(Expected := 3, Actual := AoProgress.Status.Index, Message := 'Index');
AssertEquals_DINT(Expected := 1, Actual := AoProgress.Status.RepeatsDone, Message := 'RepeatsDone');

TEST_FINISHED();
END_METHOD


METHOD PRIVATE ZeroVelocityKeepsPrevious
VAR
    Cycle : INT;
    Before : REAL;
END_VAR

TEST('ZeroVelocityKeepsPrevious');

AoZeroVelocity.Cfg.VelocityVPerS := 1.0;
AoZeroVelocity.Cfg.Setpoint := 5.0;
FOR Cycle := 1 TO 100 DO
    AoZeroVelocity();
END_FOR
Before := AoZeroVelocity.Status.Value;
AoZeroVelocity.Cfg.VelocityVPerS := 0.0;
AoZeroVelocity();
AssertTrue(Condition := AoZeroVelocity.Status.Error, Message := 'Error');
AssertTrue(Condition := FIND(AoZeroVelocity.Status.ErrorText, 'VelocityVPerS') > 0, Message := 'names the velocity');
AssertEquals_REAL(Expected := Before + 0.001, Actual := AoZeroVelocity.Status.Value, Delta := 1.0E-5, Message := 'continues at the previous velocity');

TEST_FINISHED();
END_METHOD

END_FUNCTION_BLOCK

// ---- Tests/FB_MultiTriggerTest.TcPOU

(*
    Tests of FB_MultiTrigger (specs/multi-trigger).
*)
FUNCTION_BLOCK FB_MultiTriggerTest EXTENDS TcUnit.FB_TestSuite
VAR
    TrigZero : MBIDivB.FB_MultiTrigger;
    TrigTiming : MBIDivB.FB_MultiTrigger;
    TrigTwenty : MBIDivB.FB_MultiTrigger;
    TrigContinuous : MBIDivB.FB_MultiTrigger;
    TrigSubCycle : MBIDivB.FB_MultiTrigger;
    TrigStop : MBIDivB.FB_MultiTrigger;
    TrigProgress : MBIDivB.FB_MultiTrigger;
    TrigGroup1 : MBIDivB.FB_MultiTrigger;
    TrigGroup2 : MBIDivB.FB_MultiTrigger;
    TrigGroup3 : MBIDivB.FB_MultiTrigger;
    TrigGate : MBIDivB.FB_MultiTrigger;
    CtGate : MBIDivB.FB_CounterTimer;
    TrigMethod : MBIDivB.FB_MultiTrigger;
    TrigDelayText : MBIDivB.FB_MultiTrigger;
END_VAR


ZeroCountRejected();
TimingOn1msTask();
TwentyPulses();
ContinuousUntilStop();
SubCycleHighTime();
StopDuringHigh();
ProgressAfterThirdEdge();
GroupStartEnabledOnly();
GatesCounterTimer();
MethodStartEqualsFlag();
StateTextInDelay();


METHOD PRIVATE ContinuousUntilStop
VAR
    Cycle : INT;
END_VAR

TEST('ContinuousUntilStop');

TrigContinuous.Cfg.HighMs := 1.0;
TrigContinuous.Cfg.LowMs := 1.0;
TrigContinuous.Cfg.Count := -1;
TrigContinuous.Cmd.Start := TRUE;
FOR Cycle := 1 TO 1000 DO
    TrigContinuous();
END_FOR
AssertTrue(Condition := TrigContinuous.Status.State <> 0, Message := 'still running');
AssertEquals_UDINT(Expected := 500, Actual := TrigContinuous.Status.EdgesDone, Message := 'EdgesDone');
TrigContinuous.Cmd.Stop := TRUE;
TrigContinuous();
AssertEquals_INT(Expected := 0, Actual := TrigContinuous.Status.State, Message := 'stopped');
AssertFalse(Condition := TrigContinuous.Output, Message := 'output low');

TEST_FINISHED();
END_METHOD


METHOD PRIVATE GatesCounterTimer
VAR
    Cycle : INT;
END_VAR

TEST('GatesCounterTimer');

TrigGate.Cfg.HighMs := 1.0;
TrigGate.Cfg.LowMs := 9.0;
TrigGate.Cfg.Count := 3;
CtGate.Cfg.StartMode := 1;
CtGate.Cfg.IntegrationTimeMs := 2.0;
CtGate.Cfg.Points := 3;
TrigGate.Start();
CtGate.Start();
FOR Cycle := 0 TO 30 DO   // edges in cycles 0, 10 and 20
    TrigGate();
    CtGate.Channel[1].Input := INT_TO_REAL(Cycle);
    CtGate(Gate := TrigGate.Status.Output);
END_FOR
AssertEquals_DINT(Expected := 3, Actual := CtGate.Status.PointsDone, Message := 'one point per edge');
AssertEquals_REAL(Expected := 0.5, Actual := CtGate.Channel[1].Data[1], Delta := 1.0E-6, Message := 'window 1 = cycles 0-1');
AssertEquals_REAL(Expected := 20.5, Actual := CtGate.Channel[1].Data[3], Delta := 1.0E-6, Message := 'window 3 = cycles 20-21');

TEST_FINISHED();
END_METHOD


METHOD PRIVATE GroupStartEnabledOnly
VAR
    Cycle : INT;
    Mismatch : INT;
END_VAR

TEST('GroupStartEnabledOnly');

TrigGroup1.Cfg.Enabled := TRUE;
TrigGroup2.Cfg.Enabled := TRUE;
TrigGroup3.Cfg.Enabled := FALSE;
TrigGroup1.Cfg.Count := 5;
TrigGroup2.Cfg.Count := 5;
TrigGroup3.Cfg.Count := 5;
TrigGroup1.StartIfEnabled();
TrigGroup2.StartIfEnabled();
TrigGroup3.StartIfEnabled();
FOR Cycle := 0 TO 20 DO
    TrigGroup1();
    TrigGroup2();
    TrigGroup3();
    IF TrigGroup1.Output <> TrigGroup2.Output THEN
        Mismatch := Mismatch + 1;
    END_IF
END_FOR
AssertEquals_INT(Expected := 0, Actual := Mismatch, Message := 'aligned edges');
AssertEquals_UDINT(Expected := 5, Actual := TrigGroup1.Status.EdgesDone, Message := 'trigger 1 ran');
AssertEquals_UDINT(Expected := 0, Actual := TrigGroup3.Status.EdgesDone, Message := 'disabled trigger stays idle');
AssertFalse(Condition := TrigGroup3.Status.Error, Message := 'no error on the disabled trigger');

TEST_FINISHED();
END_METHOD


METHOD PRIVATE MethodStartEqualsFlag
VAR
    Accepted : BOOL;
END_VAR

TEST('MethodStartEqualsFlag');

TrigMethod.Cfg.Count := 0;
Accepted := TrigMethod.Start();
AssertFalse(Condition := Accepted, Message := 'rejected like the flag');
AssertTrue(Condition := FIND(TrigMethod.Status.ErrorText, 'Count') > 0, Message := 'same error');
TrigMethod.Cfg.Count := 1;
TrigMethod.Cfg.DelayMs := 3.0;
Accepted := TrigMethod.Start();
AssertTrue(Condition := Accepted, Message := 'accepted');
AssertFalse(Condition := TrigMethod.Status.Error, Message := 'error cleared');
AssertEquals_INT(Expected := 1, Actual := TrigMethod.Status.State, Message := 'DELAY');

TEST_FINISHED();
END_METHOD


METHOD PRIVATE ProgressAfterThirdEdge
VAR
    Cycle : INT;
END_VAR

TEST('ProgressAfterThirdEdge');

TrigProgress.Cfg.HighMs := 2.0;
TrigProgress.Cfg.LowMs := 2.0;
TrigProgress.Cfg.Count := 10;
TrigProgress.Cmd.Start := TRUE;
FOR Cycle := 0 TO 8 DO   // edges in cycles 0, 4 and 8
    TrigProgress();
END_FOR
AssertEquals_UDINT(Expected := 3, Actual := TrigProgress.Status.EdgesDone, Message := 'EdgesDone');
AssertTrue(Condition := TrigProgress.Status.Output, Message := 'Output');
AssertEquals_INT(Expected := 2, Actual := TrigProgress.Status.State, Message := 'HIGH');

TEST_FINISHED();
END_METHOD


METHOD PRIVATE StateTextInDelay

TEST('StateTextInDelay');

TrigDelayText.Cfg.DelayMs := 5.0;
TrigDelayText.Cmd.Start := TRUE;
TrigDelayText();
AssertEquals_INT(Expected := 1, Actual := TrigDelayText.Status.State, Message := 'State');
AssertEquals_STRING(Expected := 'DELAY', Actual := TrigDelayText.Status.StateText, Message := 'StateText');

TEST_FINISHED();
END_METHOD


METHOD PRIVATE StopDuringHigh
VAR
    Cycle : INT;
END_VAR

TEST('StopDuringHigh');

TrigStop.Cfg.HighMs := 10.0;
TrigStop.Cfg.Count := 1;
TrigStop.Cmd.Start := TRUE;
FOR Cycle := 0 TO 2 DO
    TrigStop();
END_FOR
AssertTrue(Condition := TrigStop.Output, Message := 'high before the stop');
TrigStop.Cmd.Stop := TRUE;
TrigStop();
AssertFalse(Condition := TrigStop.Output, Message := 'low in the stop cycle');
AssertEquals_INT(Expected := 0, Actual := TrigStop.Status.State, Message := 'idle');

TEST_FINISHED();
END_METHOD


METHOD PRIVATE SubCycleHighTime
VAR
    Cycle : INT;
    HighCycles : INT;
END_VAR

TEST('SubCycleHighTime');

TrigSubCycle.Cfg.HighMs := 0.3;
TrigSubCycle.Cfg.LowMs := 5.0;
TrigSubCycle.Cfg.Count := 1;
TrigSubCycle.Cmd.Start := TRUE;
FOR Cycle := 0 TO 10 DO
    TrigSubCycle();
    IF TrigSubCycle.Output THEN
        HighCycles := HighCycles + 1;
    END_IF
END_FOR
AssertEquals_INT(Expected := 1, Actual := HighCycles, Message := 'one high cycle');
AssertEquals_REAL(Expected := 1.0, Actual := TrigSubCycle.Status.HighMs, Delta := 1.0E-6, Message := 'effective high time');

TEST_FINISHED();
END_METHOD


METHOD PRIVATE TimingOn1msTask
VAR
    Cycle : INT;
    Expected : BOOL;
    Wrong : INT;
END_VAR

TEST('TimingOn1msTask');

TrigTiming.Cfg.DelayMs := 5.0;
TrigTiming.Cfg.HighMs := 2.0;
TrigTiming.Cfg.LowMs := 3.0;
TrigTiming.Cfg.Count := 2;
TrigTiming.Cmd.Start := TRUE;
FOR Cycle := 0 TO 20 DO
    TrigTiming();
    Expected := Cycle = 5 OR Cycle = 6 OR Cycle = 10 OR Cycle = 11;
    IF TrigTiming.Output <> Expected THEN
        Wrong := Wrong + 1;
    END_IF
END_FOR
AssertEquals_INT(Expected := 0, Actual := Wrong, Message := 'high in cycles 5-6 and 10-11 only');
AssertEquals_INT(Expected := 0, Actual := TrigTiming.Status.State, Message := 'idle');

TEST_FINISHED();
END_METHOD


METHOD PRIVATE TwentyPulses
VAR
    Cycle : INT;
    Previous : BOOL;
    Edges : INT;
END_VAR

TEST('TwentyPulses');

TrigTwenty.Cfg.HighMs := 1.0;
TrigTwenty.Cfg.LowMs := 1.0;
TrigTwenty.Cfg.Count := 20;
TrigTwenty.Cmd.Start := TRUE;
FOR Cycle := 0 TO 100 DO
    TrigTwenty();
    IF TrigTwenty.Output AND NOT Previous THEN
        Edges := Edges + 1;
    END_IF
    Previous := TrigTwenty.Output;
END_FOR
AssertEquals_INT(Expected := 20, Actual := Edges, Message := 'exactly 20 rising edges');
AssertEquals_UDINT(Expected := 20, Actual := TrigTwenty.Status.EdgesDone, Message := 'EdgesDone');
AssertEquals_INT(Expected := 0, Actual := TrigTwenty.Status.State, Message := 'idle');

TEST_FINISHED();
END_METHOD


METHOD PRIVATE ZeroCountRejected

TEST('ZeroCountRejected');

TrigZero.Cfg.Count := 0;
TrigZero.Cmd.Start := TRUE;
TrigZero();
AssertTrue(Condition := TrigZero.Status.Error, Message := 'Error');
AssertTrue(Condition := FIND(TrigZero.Status.ErrorText, 'Count') > 0, Message := 'names Count');
AssertEquals_INT(Expected := 0, Actual := TrigZero.Status.State, Message := 'idle');

TEST_FINISHED();
END_METHOD

END_FUNCTION_BLOCK

// ---- Tests/FB_FlowMeterTest.TcPOU

(*
    Tests of FB_FlowMeter (specs/flow-meter). The overrun test needs
    FLOW_BUFFER_LENGTH < 500, because a 1 ms task produces at most 500 edges
    per second.
*)
FUNCTION_BLOCK FB_FlowMeterTest EXTENDS TcUnit.FB_TestSuite
VAR
    FlowSteady : MBIDivB.FB_FlowMeter;
    FlowOverrun : MBIDivB.FB_FlowMeter;
END_VAR


SteadyPulsesThenStop();
OverrunError();


METHOD PRIVATE OverrunError
VAR
    Cycle : INT;
END_VAR

TEST('OverrunError');

AssertTrue(Condition := MBIDivB.GVL_Param.FLOW_BUFFER_LENGTH < 500, Message := 'override FLOW_BUFFER_LENGTH below 500 in the test project');
FOR Cycle := 1 TO 1000 DO
    FlowOverrun.SensorInput := Cycle MOD 2 = 0;
    FlowOverrun();
END_FOR
AssertTrue(Condition := FlowOverrun.Status.Error, Message := 'Error');
AssertTrue(Condition := FIND(FlowOverrun.Status.ErrorText, 'out of range') > 0, Message := 'ErrorText');

TEST_FINISHED();
END_METHOD


METHOD PRIVATE SteadyPulsesThenStop
VAR
    Cycle : INT;
END_VAR

TEST('SteadyPulsesThenStop');

FOR Cycle := 1 TO 5000 DO
    FlowSteady.SensorInput := Cycle MOD 50 = 0;
    FlowSteady();
END_FOR
AssertEquals_REAL(Expected := 20.0, Actual := FlowSteady.Status.FrequencyHz, Delta := 0.0, Message := '20 Hz');
AssertEquals_REAL(Expected := 5.6, Actual := FlowSteady.Status.FlowRate, Delta := 1.0E-4, Message := 'default factor');
FlowSteady.SensorInput := FALSE;
FOR Cycle := 1 TO 1001 DO
    FlowSteady();
END_FOR
AssertEquals_REAL(Expected := 0.0, Actual := FlowSteady.Status.FrequencyHz, Delta := 0.0, Message := 'flow stopped');

TEST_FINISHED();
END_METHOD

END_FUNCTION_BLOCK

// ---- Tests/FB_ShutterControlTest.TcPOU

(*
    Tests of FB_ShutterControl (specs/shutter-control).
*)
FUNCTION_BLOCK FB_ShutterControlTest EXTENDS TcUnit.FB_TestSuite
VAR
    ShutterTable : MBIDivB.FB_ShutterControl;
    ShutterUnknown : MBIDivB.FB_ShutterControl;
    ShutterSoftware : MBIDivB.FB_ShutterControl;
    ShutterStartup : MBIDivB.FB_ShutterControl;
END_VAR


TruthTable();
UnknownModeKeepsLast();
SoftwareSwitch();
StartupState();


METHOD PRIVATE SoftwareSwitch

TEST('SoftwareSwitch');

ShutterSoftware();
ShutterSoftware.Cfg.SoftwareSignal := TRUE;
ShutterSoftware();
AssertTrue(Condition := ShutterSoftware.Output, Message := 'output in the next call');

TEST_FINISHED();
END_METHOD


METHOD PRIVATE StartupState

TEST('StartupState');

ShutterStartup.HwInput := TRUE;
ShutterStartup();
AssertFalse(Condition := ShutterStartup.Output, Message := 'output FALSE');
AssertEquals_INT(Expected := 3, Actual := ShutterStartup.Status.Mode, Message := 'mode SW');
AssertEquals_STRING(Expected := 'SW', Actual := ShutterStartup.Status.ModeText, Message := 'ModeText');

TEST_FINISHED();
END_METHOD


METHOD PRIVATE TruthTable
VAR
    Mode : INT;
    Combination : INT;
    Hw : BOOL;
    Sw : BOOL;
    Expected : BOOL;
    Wrong : INT;
END_VAR

TEST('TruthTable');

FOR Mode := 0 TO 3 DO
    FOR Combination := 0 TO 3 DO
        Hw := Combination = 1 OR Combination = 3;
        Sw := Combination = 2 OR Combination = 3;
        CASE Mode OF
            0: Expected := Hw AND Sw;
            1: Expected := Hw OR Sw;
            2: Expected := Hw;
            3: Expected := Sw;
        END_CASE
        ShutterTable.Cfg.Mode := Mode;
        ShutterTable.Cfg.SoftwareSignal := Sw;
        ShutterTable.HwInput := Hw;
        ShutterTable();
        IF ShutterTable.Output <> Expected OR ShutterTable.Status.Output <> Expected THEN
            Wrong := Wrong + 1;
        END_IF
    END_FOR
END_FOR
AssertEquals_INT(Expected := 0, Actual := Wrong, Message := 'outputs matching the mode definitions');

TEST_FINISHED();
END_METHOD


METHOD PRIVATE UnknownModeKeepsLast

TEST('UnknownModeKeepsLast');

ShutterUnknown.Cfg.Mode := 1;
ShutterUnknown();
ShutterUnknown.Cfg.Mode := 7;
ShutterUnknown.HwInput := TRUE;
ShutterUnknown.Cfg.SoftwareSignal := FALSE;
ShutterUnknown();
AssertEquals_INT(Expected := 1, Actual := ShutterUnknown.Status.Mode, Message := 'keeps OR');
AssertTrue(Condition := ShutterUnknown.Output, Message := 'OR output');
AssertTrue(Condition := ShutterUnknown.Status.Error, Message := 'Error');
AssertTrue(Condition := FIND(ShutterUnknown.Status.ErrorText, 'Mode') > 0, Message := 'names the mode');

TEST_FINISHED();
END_METHOD

END_FUNCTION_BLOCK

// ---- Tests/FB_LedControlTest.TcPOU

(*
    Tests of FB_LedControl (specs/led-control) with simulated EL2595 status
    words. Status word bits: 0 ready, 1 output active, 6 warning, 7 error.
    Control word bits: 1 output, 7 reset.
*)
FUNCTION_BLOCK FB_LedControlTest EXTENDS TcUnit.FB_TestSuite
VAR
    LedOnOff : MBIDivB.FB_LedControl;
    LedNotReady : MBIDivB.FB_LedControl;
    LedTimeout : MBIDivB.FB_LedControl;
    LedTimeout50 : MBIDivB.FB_LedControl;
    LedUnlimited : MBIDivB.FB_LedControl;
    LedNegative : MBIDivB.FB_LedControl;
    LedOnTime : MBIDivB.FB_LedControl;
    LedCurrent : MBIDivB.FB_LedControl;
    LedRange : MBIDivB.FB_LedControl;
    LedReadback : MBIDivB.FB_LedControl;
    LedFault : MBIDivB.FB_LedControl;
    LedReset : MBIDivB.FB_LedControl;
END_VAR


SwitchOnAndOff();
NotReadyRejected();
Timeout500ms();
Timeout50ms();
UnlimitedOnTime();
NegativeMaxOnTimeRejected();
OnTimeDisplayed();
CurrentChangeWhileOn();
CurrentOutOfRange();
VoltageAndCurrentReadback();
TerminalErrorToFault();
ResetPulseOneCycle();


METHOD PRIVATE CurrentChangeWhileOn

TEST('CurrentChangeWhileOn');

LedCurrent.StatusWord := 16#0001;
LedCurrent.Cfg.CurrentMa := 400;
LedCurrent.Cmd.On := TRUE;
LedCurrent();
AssertEquals_UINT(Expected := 400, Actual := LedCurrent.CurrentSetpoint, Message := '400 mA');
LedCurrent.Cfg.CurrentMa := 500;
LedCurrent();
AssertEquals_UINT(Expected := 500, Actual := LedCurrent.CurrentSetpoint, Message := '500 mA in the next cycle');
AssertEquals_INT(Expected := 1, Actual := LedCurrent.Status.State, Message := 'still on');

TEST_FINISHED();
END_METHOD


METHOD PRIVATE CurrentOutOfRange

TEST('CurrentOutOfRange');

LedRange.Cfg.CurrentMa := 400;
LedRange();
LedRange.Cfg.CurrentMa := 1000;
LedRange();
AssertEquals_UINT(Expected := 400, Actual := LedRange.CurrentSetpoint, Message := 'last valid value kept');
AssertTrue(Condition := FIND(LedRange.Status.ErrorText, 'CurrentMa') > 0, Message := 'names CurrentMa');

TEST_FINISHED();
END_METHOD


METHOD PRIVATE NegativeMaxOnTimeRejected

TEST('NegativeMaxOnTimeRejected');

LedNegative.StatusWord := 16#0001;
LedNegative.Cfg.MaxOnTimeMs := -1.0;
LedNegative.Cmd.On := TRUE;
LedNegative();
AssertEquals_INT(Expected := 0, Actual := LedNegative.Status.State, Message := 'stays off');
AssertTrue(Condition := FIND(LedNegative.Status.ErrorText, 'MaxOnTimeMs') > 0, Message := 'names MaxOnTimeMs');

TEST_FINISHED();
END_METHOD


METHOD PRIVATE NotReadyRejected

TEST('NotReadyRejected');

LedNotReady.StatusWord := 16#0000;
LedNotReady.Cmd.On := TRUE;
LedNotReady();
AssertTrue(Condition := (LedNotReady.ControlWord AND 16#0002) = 0, Message := 'stays off');
AssertTrue(Condition := LedNotReady.Status.Error, Message := 'Error');
AssertTrue(Condition := FIND(LedNotReady.Status.ErrorText, 'not ready') > 0, Message := 'ErrorText');

TEST_FINISHED();
END_METHOD


METHOD PRIVATE OnTimeDisplayed
VAR
    Cycle : INT;
END_VAR

TEST('OnTimeDisplayed');

LedOnTime.StatusWord := 16#0001;
LedOnTime.Cmd.On := TRUE;
FOR Cycle := 1 TO 200 DO
    LedOnTime();
END_FOR
AssertEquals_REAL(Expected := 200.0, Actual := LedOnTime.Status.OnTimeMs, Delta := 1.0, Message := 'OnTimeMs while on');
LedOnTime.Cmd.On := TRUE;   // accepted without restarting the on time
LedOnTime();
AssertEquals_REAL(Expected := 201.0, Actual := LedOnTime.Status.OnTimeMs, Delta := 1.0, Message := 'On while on keeps the on time');
LedOnTime.Cmd.Off := TRUE;
FOR Cycle := 1 TO 50 DO
    LedOnTime();
END_FOR
AssertEquals_REAL(Expected := 201.0, Actual := LedOnTime.Status.OnTimeMs, Delta := 1.0, Message := 'last on period while off');

TEST_FINISHED();
END_METHOD


METHOD PRIVATE ResetPulseOneCycle

TEST('ResetPulseOneCycle');

LedReset.Cmd.Reset := TRUE;
LedReset();
AssertTrue(Condition := (LedReset.ControlWord AND 16#0080) <> 0, Message := 'reset bit set');
LedReset();
AssertTrue(Condition := (LedReset.ControlWord AND 16#0080) = 0, Message := 'reset bit cleared after one cycle');

TEST_FINISHED();
END_METHOD


METHOD PRIVATE SwitchOnAndOff

TEST('SwitchOnAndOff');

LedOnOff();
AssertEquals_INT(Expected := 0, Actual := LedOnOff.Status.State, Message := 'off after start');
LedOnOff.StatusWord := 16#0001;
LedOnOff.Cmd.On := TRUE;
LedOnOff();
AssertTrue(Condition := (LedOnOff.ControlWord AND 16#0002) <> 0, Message := 'output bit set');
AssertEquals_STRING(Expected := 'ON', Actual := LedOnOff.Status.StateText, Message := 'ON');
LedOnOff.Cmd.Off := TRUE;
LedOnOff();
AssertTrue(Condition := (LedOnOff.ControlWord AND 16#0002) = 0, Message := 'output bit cleared');
AssertEquals_STRING(Expected := 'OFF', Actual := LedOnOff.Status.StateText, Message := 'OFF');

TEST_FINISHED();
END_METHOD


METHOD PRIVATE TerminalErrorToFault

TEST('TerminalErrorToFault');

LedFault.StatusWord := 16#0001;
LedFault.Cmd.On := TRUE;
LedFault();
LedFault.StatusWord := 16#0081;
LedFault();
AssertTrue(Condition := (LedFault.ControlWord AND 16#0002) = 0, Message := 'output deactivated');
AssertEquals_STRING(Expected := 'FAULT', Actual := LedFault.Status.StateText, Message := 'FAULT');
AssertTrue(Condition := LedFault.Status.Error, Message := 'Error');
AssertTrue(Condition := FIND(LedFault.Status.ErrorText, '0xA000') > 0, Message := 'refers to the diag data');

TEST_FINISHED();
END_METHOD


METHOD PRIVATE Timeout500ms
VAR
    Cycle : INT;
    OnCycles : INT;
END_VAR

TEST('Timeout500ms');

LedTimeout.StatusWord := 16#0001;
LedTimeout.Cfg.MaxOnTimeMs := 500.0;
LedTimeout.Cmd.On := TRUE;
FOR Cycle := 1 TO 600 DO
    LedTimeout();
    IF (LedTimeout.ControlWord AND 16#0002) <> 0 THEN
        OnCycles := OnCycles + 1;
    END_IF
END_FOR
AssertEquals_INT(Expected := 500, Actual := OnCycles, Message := 'on for 500 cycles');
AssertEquals_STRING(Expected := 'TIMEOUT', Actual := LedTimeout.Status.StateText, Message := 'TIMEOUT');

TEST_FINISHED();
END_METHOD


METHOD PRIVATE Timeout50ms
VAR
    Cycle : INT;
    OnCycles : INT;
END_VAR

TEST('Timeout50ms');

LedTimeout50.StatusWord := 16#0001;
LedTimeout50.Cfg.MaxOnTimeMs := 50.0;
LedTimeout50.Cmd.On := TRUE;
FOR Cycle := 1 TO 100 DO
    LedTimeout50();
    IF (LedTimeout50.ControlWord AND 16#0002) <> 0 THEN
        OnCycles := OnCycles + 1;
    END_IF
END_FOR
AssertEquals_INT(Expected := 50, Actual := OnCycles, Message := 'deactivated after 50 cycles');
AssertEquals_INT(Expected := 2, Actual := LedTimeout50.Status.State, Message := 'TIMEOUT');

TEST_FINISHED();
END_METHOD


METHOD PRIVATE UnlimitedOnTime
VAR
    Cycle : INT;
END_VAR

TEST('UnlimitedOnTime');

LedUnlimited.StatusWord := 16#0001;
LedUnlimited.Cfg.MaxOnTimeMs := 0.0;
LedUnlimited.Cmd.On := TRUE;
FOR Cycle := 1 TO 10000 DO
    LedUnlimited();
END_FOR
AssertEquals_INT(Expected := 1, Actual := LedUnlimited.Status.State, Message := 'still on');
LedUnlimited.Cmd.Off := TRUE;
LedUnlimited();
AssertEquals_INT(Expected := 0, Actual := LedUnlimited.Status.State, Message := 'off');

TEST_FINISHED();
END_METHOD


METHOD PRIVATE VoltageAndCurrentReadback

TEST('VoltageAndCurrentReadback');

LedReadback.InfoData1 := 1230;
LedReadback.InfoData2 := 500;
LedReadback();
AssertEquals_REAL(Expected := 12.3, Actual := LedReadback.Status.VoltageV, Delta := 1.0E-4, Message := 'VoltageV');
AssertEquals_REAL(Expected := 500.0, Actual := LedReadback.Status.CurrentMa, Delta := 1.0E-4, Message := 'CurrentMa');

TEST_FINISHED();
END_METHOD

END_FUNCTION_BLOCK

// ---- Tests/FB_FemtoAmplifierTest.TcPOU

(*
    Tests of FB_FemtoAmplifier (specs/femto-amplifier). Settling times
    assume the 1 ms test task: 150 ms = 150 calls.

    AiShared is never called; it only gives the blocks that do not test the
    current an assigned input, so that no input error hides the result.
*)
FUNCTION_BLOCK FB_FemtoAmplifierTest EXTENDS TcUnit.FB_TestSuite
VAR
    AiShared : MBIDivB.FB_AnalogInput16;
    FemtoLowest : MBIDivB.FB_FemtoAmplifier;
    FemtoHighest : MBIDivB.FB_FemtoAmplifier;
    FemtoTable : MBIDivB.FB_FemtoAmplifier;
    FemtoModeSwitch : MBIDivB.FB_FemtoAmplifier;
    FemtoRange : MBIDivB.FB_FemtoAmplifier;
    FemtoReadback : MBIDivB.FB_FemtoAmplifier;
    FemtoAc : MBIDivB.FB_FemtoAmplifier;
    FemtoSettling : MBIDivB.FB_FemtoAmplifier;
    FemtoChange : MBIDivB.FB_FemtoAmplifier;
    FemtoTimeChange : MBIDivB.FB_FemtoAmplifier;
    FemtoZero : MBIDivB.FB_FemtoAmplifier;
    FemtoNegativeTime : MBIDivB.FB_FemtoAmplifier;
    FemtoOverload : MBIDivB.FB_FemtoAmplifier;
    AiCurrent : MBIDivB.FB_AnalogInput16;
    FemtoCurrent : MBIDivB.FB_FemtoAmplifier;
    AiNegative : MBIDivB.FB_AnalogInput32;
    FemtoNegative : MBIDivB.FB_FemtoAmplifier;
    AiMixing : MBIDivB.FB_AnalogInput16;
    FemtoMixing : MBIDivB.FB_FemtoAmplifier;
    FemtoMissing : MBIDivB.FB_FemtoAmplifier;
    FemtoStartup : MBIDivB.FB_FemtoAmplifier;
END_VAR


LowestLowNoiseGain();
HighestHighSpeedGain();
BitTable();
ModeSwitchedBeforeExponent();
ExponentOutOfRange();
GainReadback();
AcCoupling();
DefaultSettling();
ChangeDuringSettling();
SettlingTimeChangedDuringSettling();
ZeroSettlingTime();
NegativeSettlingTime();
OverloadNoError();
CurrentFromVoltage();
NegativeCurrent();
NoMixingOfGains();
MissingInput();
StartupState();


METHOD PRIVATE AcCoupling

TEST('AcCoupling');

FemtoAc(Input := AiShared);
AssertTrue(Condition := FemtoAc.DcCoupling, Message := 'DC after start');
FemtoAc.Cfg.DcCoupling := FALSE;
FemtoAc();
AssertFalse(Condition := FemtoAc.DcCoupling, Message := 'AC output in the next call');
AssertFalse(Condition := FemtoAc.Status.DcCoupling, Message := 'Status.DcCoupling');

TEST_FINISHED();
END_METHOD


METHOD PRIVATE BitTable
VAR
    Mode : INT;
    LowNoise : BOOL;
    FirstExponent : INT;
    Exponent : INT;
    Code : INT;
    Wrong : INT;
    Code7 : INT;
END_VAR

TEST('BitTable');

// DLPCA-200 table: code 0 is 10^3 V/A low noise or 10^5 V/A high speed.
FOR Mode := 0 TO 1 DO
    LowNoise := Mode = 0;
    IF LowNoise THEN
        FirstExponent := 3;
    ELSE
        FirstExponent := 5;
    END_IF
    FOR Exponent := FirstExponent TO FirstExponent + 6 DO
        FemtoTable.Cfg.LowNoise := LowNoise;
        FemtoTable.Cfg.GainExponent := Exponent;
        FemtoTable(Input := AiShared);
        Code := OutputCode(Femto := FemtoTable);
        IF Code <> Exponent - FirstExponent OR FemtoTable.LowNoise <> LowNoise OR FemtoTable.Status.Error THEN
            Wrong := Wrong + 1;
        END_IF
        IF Code = 7 THEN
            Code7 := Code7 + 1;
        END_IF
    END_FOR
END_FOR
AssertEquals_INT(Expected := 0, Actual := Wrong, Message := 'settings not matching the bit table');
AssertEquals_INT(Expected := 0, Actual := Code7, Message := 'code 7 output');

TEST_FINISHED();
END_METHOD


METHOD PRIVATE ChangeDuringSettling
VAR
    Call : INT;
END_VAR

TEST('ChangeDuringSettling');

FemtoChange(Input := AiShared);
CountSettlingCalls(Femto := FemtoChange);
FemtoChange.Cfg.GainExponent := 4;
FOR Call := 1 TO 100 DO
    FemtoChange();
END_FOR
FemtoChange.Cfg.GainExponent := 5;
AssertEquals_INT(Expected := 150, Actual := CountSettlingCalls(Femto := FemtoChange), Message := 'SETTLING calls after the second change');

TEST_FINISHED();
END_METHOD


(*
    Calls Femto until it reports READY and returns the number of calls that
    reported SETTLING. Stops after 1000 calls.
*)
METHOD PRIVATE CountSettlingCalls : INT
VAR_IN_OUT
    Femto : MBIDivB.FB_FemtoAmplifier;
END_VAR
VAR
    Call : INT;
END_VAR

CountSettlingCalls := 0;
FOR Call := 1 TO 1000 DO
    Femto();
    IF Femto.Status.State <> 1 THEN
        RETURN;
    END_IF
    CountSettlingCalls := CountSettlingCalls + 1;
END_FOR
END_METHOD


METHOD PRIVATE CurrentFromVoltage

TEST('CurrentFromVoltage');

AiCurrent.SetScale(RawFullScale := 1000, ValueFullScale := 1.0);
AiCurrent.Raw := 2000;
FemtoCurrent.Cfg.GainExponent := 6;
AiCurrent();
FemtoCurrent(Input := AiCurrent);
AssertEquals_REAL(Expected := 2.0E-6, Actual := FemtoCurrent.Status.CurrentA, Delta := 1.0E-12, Message := 'CurrentA');
AssertFalse(Condition := FemtoCurrent.Status.Error, Message := 'Error');

TEST_FINISHED();
END_METHOD


METHOD PRIVATE DefaultSettling

TEST('DefaultSettling');

FemtoSettling(Input := AiShared);
CountSettlingCalls(Femto := FemtoSettling);
FemtoSettling.Cfg.GainExponent := 4;
AssertEquals_INT(Expected := 150, Actual := CountSettlingCalls(Femto := FemtoSettling), Message := 'SETTLING calls');
AssertEquals_INT(Expected := 0, Actual := FemtoSettling.Status.State, Message := 'READY afterwards');
AssertFalse(Condition := FemtoSettling.Status.Settling, Message := 'Status.Settling afterwards');

TEST_FINISHED();
END_METHOD


METHOD PRIVATE ExponentOutOfRange

TEST('ExponentOutOfRange');

FemtoRange.Cfg.LowNoise := FALSE;
FemtoRange.Cfg.GainExponent := 7;
FemtoRange(Input := AiShared);
FemtoRange.Cfg.GainExponent := 12;
FemtoRange();
AssertEquals_INT(Expected := 7, Actual := FemtoRange.Status.GainExponent, Message := 'last valid gain in use');
AssertEquals_INT(Expected := 2, Actual := OutputCode(Femto := FemtoRange), Message := 'outputs keep 10^7 V/A');
AssertTrue(Condition := FemtoRange.Status.Error, Message := 'Error');
AssertTrue(Condition := FIND(FemtoRange.Status.ErrorText, 'GainExponent') > 0, Message := 'names GainExponent');
AssertTrue(Condition := FIND(FemtoRange.Status.ErrorText, '5..11') > 0, Message := 'names the valid range');

TEST_FINISHED();
END_METHOD


METHOD PRIVATE GainReadback

TEST('GainReadback');

FemtoReadback.Cfg.GainExponent := 7;
FemtoReadback(Input := AiShared);
AssertEquals_REAL(Expected := 1.0E7, Actual := FemtoReadback.Status.GainVPerA, Delta := 0.5, Message := 'GainVPerA');
AssertEquals_INT(Expected := 7, Actual := FemtoReadback.Status.GainExponent, Message := 'GainExponent');

TEST_FINISHED();
END_METHOD


METHOD PRIVATE HighestHighSpeedGain

TEST('HighestHighSpeedGain');

FemtoHighest.Cfg.LowNoise := FALSE;
FemtoHighest.Cfg.GainExponent := 11;
FemtoHighest(Input := AiShared);
AssertTrue(Condition := FemtoHighest.GainBit2, Message := 'pin 12');
AssertTrue(Condition := FemtoHighest.GainBit1, Message := 'pin 11');
AssertFalse(Condition := FemtoHighest.GainBit0, Message := 'pin 10');
AssertFalse(Condition := FemtoHighest.LowNoise, Message := 'pin 14 high speed');

TEST_FINISHED();
END_METHOD


METHOD PRIVATE LowestLowNoiseGain

TEST('LowestLowNoiseGain');

FemtoLowest.Cfg.LowNoise := TRUE;
FemtoLowest.Cfg.GainExponent := 3;
FemtoLowest(Input := AiShared);
AssertFalse(Condition := FemtoLowest.GainBit2, Message := 'pin 12');
AssertFalse(Condition := FemtoLowest.GainBit1, Message := 'pin 11');
AssertFalse(Condition := FemtoLowest.GainBit0, Message := 'pin 10');
AssertTrue(Condition := FemtoLowest.LowNoise, Message := 'pin 14 low noise');

TEST_FINISHED();
END_METHOD


METHOD PRIVATE MissingInput

TEST('MissingInput');

FemtoMissing();
AssertTrue(Condition := FemtoMissing.Status.Error, Message := 'Error');
AssertTrue(Condition := FIND(FemtoMissing.Status.ErrorText, 'Input') > 0, Message := 'names the input');
AssertEquals_REAL(Expected := 0.0, Actual := FemtoMissing.Status.CurrentA, Delta := 0.0, Message := 'CurrentA');
AssertEquals_REAL(Expected := 0.0, Actual := FemtoMissing.Status.CurrentFilteredA, Delta := 0.0, Message := 'CurrentFilteredA');
FemtoMissing.Cfg.GainExponent := 5;
FemtoMissing();
AssertEquals_INT(Expected := 5, Actual := FemtoMissing.Status.GainExponent, Message := 'gain change applied');
AssertEquals_INT(Expected := 2, Actual := OutputCode(Femto := FemtoMissing), Message := 'outputs select 10^5 V/A low noise');

TEST_FINISHED();
END_METHOD


METHOD PRIVATE ModeSwitchedBeforeExponent

TEST('ModeSwitchedBeforeExponent');

FemtoModeSwitch(Input := AiShared);
FemtoModeSwitch.Cfg.LowNoise := FALSE;
FemtoModeSwitch();
AssertTrue(Condition := FemtoModeSwitch.Status.Error, Message := 'Error after the first write');
AssertEquals_INT(Expected := 0, Actual := OutputCode(Femto := FemtoModeSwitch), Message := 'still 10^3 V/A');
AssertTrue(Condition := FemtoModeSwitch.LowNoise, Message := 'still low noise');
FemtoModeSwitch.Cfg.GainExponent := 5;
FemtoModeSwitch();
AssertFalse(Condition := FemtoModeSwitch.Status.Error, Message := 'Error after the second write');
AssertEquals_INT(Expected := 0, Actual := OutputCode(Femto := FemtoModeSwitch), Message := 'code of 10^5 V/A high speed');
AssertFalse(Condition := FemtoModeSwitch.LowNoise, Message := 'high speed');
AssertEquals_INT(Expected := 5, Actual := FemtoModeSwitch.Status.GainExponent, Message := 'GainExponent');

TEST_FINISHED();
END_METHOD


METHOD PRIVATE NegativeCurrent

TEST('NegativeCurrent');

AiNegative.SetScale(RawFullScale := 1000, ValueFullScale := 1.0);
AiNegative.Raw := -500;
FemtoNegative.Cfg.GainExponent := 9;
AiNegative();
FemtoNegative(Input := AiNegative);
AssertEquals_REAL(Expected := -5.0E-10, Actual := FemtoNegative.Status.CurrentA, Delta := 1.0E-16, Message := 'CurrentA');

TEST_FINISHED();
END_METHOD


METHOD PRIVATE NegativeSettlingTime

TEST('NegativeSettlingTime');

FemtoNegativeTime(Input := AiShared);
FemtoNegativeTime.Cfg.SettlingTimeMs := -1.0;
FemtoNegativeTime();
AssertTrue(Condition := FemtoNegativeTime.Status.Error, Message := 'Error');
AssertTrue(Condition := FIND(FemtoNegativeTime.Status.ErrorText, 'SettlingTimeMs') > 0, Message := 'names SettlingTimeMs');
AssertEquals_REAL(Expected := 150.0, Actual := FemtoNegativeTime.Status.SettlingTimeMs, Delta := 1.0E-3, Message := 'previous value kept');

TEST_FINISHED();
END_METHOD


METHOD PRIVATE NoMixingOfGains
VAR
    Call : INT;
    Wrong : INT;
END_VAR

TEST('NoMixingOfGains');

AiMixing.SetScale(RawFullScale := 1000, ValueFullScale := 1.0);
AiMixing.Cfg.FilterSize := 100;
FemtoMixing.Cfg.GainExponent := 5;
FemtoMixing.Cfg.SettlingTimeMs := 10.0;

// 1.0 V at 10^5 V/A until settled and the average is full
AiMixing.Raw := 1000;
FOR Call := 1 TO 200 DO
    AiMixing();
    FemtoMixing(Input := AiMixing);
END_FOR
AssertEquals_REAL(Expected := 1.0E-5, Actual := FemtoMixing.Status.CurrentFilteredA, Delta := 1.0E-11, Message := 'filtered at 10^5 V/A');

// Gain change to 10^6 V/A; while settling the output moves to 2.0 V.
// The filtered current must equal the current until settling has ended.
FemtoMixing.Cfg.GainExponent := 6;
AiMixing.Raw := 2000;
FOR Call := 1 TO 100 DO
    AiMixing();
    FemtoMixing();
    IF FemtoMixing.Status.CurrentFilteredA <> FemtoMixing.Status.CurrentA THEN
        Wrong := Wrong + 1;
    END_IF
    IF FemtoMixing.Status.State = 0 THEN
        EXIT;
    END_IF
END_FOR
AssertEquals_INT(Expected := 0, Actual := FemtoMixing.Status.State, Message := 'READY after settling');
AssertEquals_INT(Expected := 0, Actual := Wrong, Message := 'calls with CurrentFilteredA <> CurrentA while settling');

// After settling ended, only new voltages count.
AiMixing.Raw := 3000;
FOR Call := 1 TO 5 DO
    AiMixing();
    FemtoMixing();
    IF ABS(FemtoMixing.Status.CurrentFilteredA - 3.0E-6) > 1.0E-12 THEN
        Wrong := Wrong + 1;
    END_IF
END_FOR
AssertEquals_INT(Expected := 0, Actual := Wrong, Message := 'calls with CurrentFilteredA <> 3.0E-6 A after settling');

TEST_FINISHED();
END_METHOD


(*
    Gain code on the three gain outputs of Femto: pin 12 MSB, pin 10 LSB.
*)
METHOD PRIVATE OutputCode : INT
VAR_IN_OUT
    Femto : MBIDivB.FB_FemtoAmplifier;
END_VAR

OutputCode := 4 * BOOL_TO_INT(Femto.GainBit2) + 2 * BOOL_TO_INT(Femto.GainBit1) + BOOL_TO_INT(Femto.GainBit0);
END_METHOD


METHOD PRIVATE OverloadNoError

TEST('OverloadNoError');

FemtoOverload(Input := AiShared);
FemtoOverload.Overload := TRUE;
FemtoOverload();
AssertTrue(Condition := FemtoOverload.Status.Overload, Message := 'Status.Overload');
AssertFalse(Condition := FemtoOverload.Status.Error, Message := 'Error');

TEST_FINISHED();
END_METHOD


METHOD PRIVATE SettlingTimeChangedDuringSettling
VAR
    Call : INT;
END_VAR

TEST('SettlingTimeChangedDuringSettling');

FemtoTimeChange(Input := AiShared);
CountSettlingCalls(Femto := FemtoTimeChange);
FemtoTimeChange.Cfg.GainExponent := 4;
FOR Call := 1 TO 20 DO
    FemtoTimeChange();
END_FOR
FemtoTimeChange.Cfg.SettlingTimeMs := 10.0;
AssertEquals_INT(Expected := 130, Actual := CountSettlingCalls(Femto := FemtoTimeChange), Message := 'remaining SETTLING calls of the running period');
AssertEquals_REAL(Expected := 10.0, Actual := FemtoTimeChange.Status.SettlingTimeMs, Delta := 1.0E-3, Message := 'Status.SettlingTimeMs');
FemtoTimeChange.Cfg.GainExponent := 5;
AssertEquals_INT(Expected := 10, Actual := CountSettlingCalls(Femto := FemtoTimeChange), Message := 'SETTLING calls of the next period');

TEST_FINISHED();
END_METHOD


METHOD PRIVATE StartupState

TEST('StartupState');

FemtoStartup(Input := AiShared);
AssertEquals_INT(Expected := 0, Actual := OutputCode(Femto := FemtoStartup), Message := 'code of 10^3 V/A');
AssertTrue(Condition := FemtoStartup.LowNoise, Message := 'low noise');
AssertTrue(Condition := FemtoStartup.DcCoupling, Message := 'DC coupling');
AssertEquals_INT(Expected := 1, Actual := FemtoStartup.Status.State, Message := 'State');
AssertEquals_STRING(Expected := 'SETTLING', Actual := FemtoStartup.Status.StateText, Message := 'StateText');
AssertTrue(Condition := FemtoStartup.Status.Settling, Message := 'Status.Settling');
AssertEquals_REAL(Expected := 150.0, Actual := FemtoStartup.Status.SettlingTimeMs, Delta := 1.0E-3, Message := 'SettlingTimeMs');
AssertEquals_REAL(Expected := 1.0E3, Actual := FemtoStartup.Status.GainVPerA, Delta := 1.0E-3, Message := 'GainVPerA');

TEST_FINISHED();
END_METHOD


METHOD PRIVATE ZeroSettlingTime

TEST('ZeroSettlingTime');

FemtoZero(Input := AiShared);
CountSettlingCalls(Femto := FemtoZero);
FemtoZero.Cfg.SettlingTimeMs := 0.0;
FemtoZero.Cfg.GainExponent := 4;
FemtoZero();
AssertEquals_INT(Expected := 0, Actual := FemtoZero.Status.State, Message := 'READY in the call of the change');

TEST_FINISHED();
END_METHOD

END_FUNCTION_BLOCK

// ---- Tests/FB_EndPositionSwitchesTest.TcPOU

(*
    Tests of FB_EndPositionSwitches (specs/end-position-switches).
*)
FUNCTION_BLOCK FB_EndPositionSwitchesTest EXTENDS TcUnit.FB_TestSuite
VAR
    ValveTable : MBIDivB.FB_EndPositionSwitches;
    ValveNeither : MBIDivB.FB_EndPositionSwitches;
    ValveFault : MBIDivB.FB_EndPositionSwitches;
END_VAR


AllCombinations();
NeitherActiveNoError();
WiringFaultClears();


METHOD PRIVATE AllCombinations
VAR
    Combination : INT;
    Open : BOOL;
    Closed : BOOL;
    ExpectedText : STRING(20);
    Wrong : INT;
END_VAR

TEST('AllCombinations');

FOR Combination := 0 TO 3 DO
    Open := Combination = 1 OR Combination = 3;
    Closed := Combination = 2 OR Combination = 3;
    CASE Combination OF
        0: ExpectedText := 'BETWEEN';
        1: ExpectedText := 'OPEN';
        2: ExpectedText := 'CLOSED';
        3: ExpectedText := 'FAULT';
    END_CASE
    ValveTable.OpenSwitch := Open;
    ValveTable.ClosedSwitch := Closed;
    ValveTable();
    IF ValveTable.Status.State <> Combination
        OR ValveTable.Status.StateText <> ExpectedText
        OR ValveTable.Status.Error <> (Combination = 3)
        OR ValveTable.Status.OpenSwitch <> Open
        OR ValveTable.Status.ClosedSwitch <> Closed
    THEN
        Wrong := Wrong + 1;
    END_IF
END_FOR
AssertEquals_INT(Expected := 0, Actual := Wrong, Message := 'combinations with a wrong state, text, error or readback');

TEST_FINISHED();
END_METHOD


METHOD PRIVATE NeitherActiveNoError
VAR
    Call : INT;
END_VAR

TEST('NeitherActiveNoError');

FOR Call := 1 TO 10000 DO
    ValveNeither();
END_FOR
AssertEquals_INT(Expected := 0, Actual := ValveNeither.Status.State, Message := 'State');
AssertEquals_STRING(Expected := 'BETWEEN', Actual := ValveNeither.Status.StateText, Message := 'StateText');
AssertFalse(Condition := ValveNeither.Status.Error, Message := 'no timeout error');

TEST_FINISHED();
END_METHOD


METHOD PRIVATE WiringFaultClears

TEST('WiringFaultClears');

ValveFault.OpenSwitch := TRUE;
ValveFault.ClosedSwitch := TRUE;
ValveFault();
AssertTrue(Condition := ValveFault.Status.Error, Message := 'Error while both are active');
AssertTrue(Condition := FIND(ValveFault.Status.ErrorText, 'Both end-position switches') > 0, Message := 'ErrorText');
ValveFault.ClosedSwitch := FALSE;
ValveFault();
AssertFalse(Condition := ValveFault.Status.Error, Message := 'Error cleared');
AssertEquals_STRING(Expected := '', Actual := ValveFault.Status.ErrorText, Message := 'ErrorText cleared');
AssertEquals_STRING(Expected := 'OPEN', Actual := ValveFault.Status.StateText, Message := 'OPEN afterwards');

TEST_FINISHED();
END_METHOD

END_FUNCTION_BLOCK

// ---- Tests/FB_PlcShutdownTest.TcPOU

(*
    Tests of FB_PlcShutdown (specs/plc-shutdown). Only FB_PlcShutdownTestable
    is used, so no request reaches the operating system of the test PC.
*)
FUNCTION_BLOCK FB_PlcShutdownTest EXTENDS TcUnit.FB_TestSuite
VAR
    ShutdownHandshake : FB_PlcShutdownTestable;
    ShutdownMethod : FB_PlcShutdownTestable;
    ShutdownRounded : FB_PlcShutdownTestable;
    ShutdownNegative : FB_PlcShutdownTestable;
    ShutdownSecond : FB_PlcShutdownTestable;
    ShutdownFails : FB_PlcShutdownTestable;
END_VAR


CommandHandshake();
ShutdownMethodAccepted();
DelayRounded();
NegativeDelayRejected();
SecondCommandRejected();
RequestFails();


METHOD PRIVATE CommandHandshake

TEST('CommandHandshake');

ShutdownHandshake.BusyCalls := 2;
ShutdownHandshake.Cmd.Shutdown := TRUE;
ShutdownHandshake();
AssertFalse(Condition := ShutdownHandshake.Cmd.Shutdown, Message := 'flag cleared');
AssertEquals_INT(Expected := 1, Actual := ShutdownHandshake.Status.State, Message := 'REQUESTING while busy');
AssertEquals_INT(Expected := 1, Actual := ShutdownHandshake.Requests, Message := 'one request sent');
AssertEquals_UDINT(Expected := 3, Actual := ShutdownHandshake.LastDelayS, Message := 'delay 3 s');
AssertEquals_REAL(Expected := 3000.0, Actual := ShutdownHandshake.Status.DelayMs, Delta := 1.0E-3, Message := 'Status.DelayMs');
ShutdownHandshake();
AssertEquals_INT(Expected := 1, Actual := ShutdownHandshake.Status.State, Message := 'REQUESTING in the second busy call');
ShutdownHandshake();
AssertEquals_INT(Expected := 2, Actual := ShutdownHandshake.Status.State, Message := 'SHUTTING_DOWN once accepted');
AssertEquals_STRING(Expected := 'SHUTTING_DOWN', Actual := ShutdownHandshake.Status.StateText, Message := 'StateText');
AssertFalse(Condition := ShutdownHandshake.Status.Error, Message := 'Error');
AssertEquals_INT(Expected := 1, Actual := ShutdownHandshake.Requests, Message := 'still one request');

TEST_FINISHED();
END_METHOD


METHOD PRIVATE DelayRounded

TEST('DelayRounded');

ShutdownRounded.Cfg.DelayMs := 2400.0;
ShutdownRounded.Cmd.Shutdown := TRUE;
ShutdownRounded();
AssertEquals_REAL(Expected := 2000.0, Actual := ShutdownRounded.Status.DelayMs, Delta := 1.0E-3, Message := 'Status.DelayMs');
AssertEquals_UDINT(Expected := 2, Actual := ShutdownRounded.LastDelayS, Message := 'request delay in s');

TEST_FINISHED();
END_METHOD


METHOD PRIVATE NegativeDelayRejected

TEST('NegativeDelayRejected');

ShutdownNegative.Cfg.DelayMs := -1.0;
ShutdownNegative.Cmd.Shutdown := TRUE;
ShutdownNegative();
AssertFalse(Condition := ShutdownNegative.Cmd.Shutdown, Message := 'flag cleared');
AssertEquals_INT(Expected := 0, Actual := ShutdownNegative.Status.State, Message := 'stays IDLE');
AssertTrue(Condition := ShutdownNegative.Status.Error, Message := 'Error');
AssertTrue(Condition := FIND(ShutdownNegative.Status.ErrorText, 'DelayMs') > 0, Message := 'names DelayMs');
AssertEquals_INT(Expected := 0, Actual := ShutdownNegative.Requests, Message := 'no request sent');

TEST_FINISHED();
END_METHOD


METHOD PRIVATE RequestFails

TEST('RequestFails');

ShutdownFails.BusyCalls := 1;
ShutdownFails.Fail := TRUE;
ShutdownFails.FailErrorId := 1793;
ShutdownFails.Cmd.Shutdown := TRUE;
ShutdownFails();
ShutdownFails();
AssertEquals_INT(Expected := 0, Actual := ShutdownFails.Status.State, Message := 'back to IDLE');
AssertTrue(Condition := ShutdownFails.Status.Error, Message := 'Error');
AssertTrue(Condition := FIND(ShutdownFails.Status.ErrorText, '1793') > 0, Message := 'ErrorText contains the error code');

// A later command sends a new request.
ShutdownFails.Fail := FALSE;
ShutdownFails.Cmd.Shutdown := TRUE;
ShutdownFails();
ShutdownFails();
AssertEquals_INT(Expected := 2, Actual := ShutdownFails.Requests, Message := 'second request sent');
AssertEquals_INT(Expected := 2, Actual := ShutdownFails.Status.State, Message := 'SHUTTING_DOWN after the retry');
AssertFalse(Condition := ShutdownFails.Status.Error, Message := 'accepted command clears the error');

TEST_FINISHED();
END_METHOD


METHOD PRIVATE SecondCommandRejected

TEST('SecondCommandRejected');

ShutdownSecond.BusyCalls := 0;
ShutdownSecond.Cmd.Shutdown := TRUE;
ShutdownSecond();
AssertEquals_INT(Expected := 2, Actual := ShutdownSecond.Status.State, Message := 'SHUTTING_DOWN');
ShutdownSecond.Cmd.Shutdown := TRUE;
ShutdownSecond();
AssertFalse(Condition := ShutdownSecond.Cmd.Shutdown, Message := 'flag cleared');
AssertEquals_INT(Expected := 2, Actual := ShutdownSecond.Status.State, Message := 'stays SHUTTING_DOWN');
AssertTrue(Condition := ShutdownSecond.Status.Error, Message := 'rejected');
AssertEquals_INT(Expected := 1, Actual := ShutdownSecond.Requests, Message := 'no second request');

TEST_FINISHED();
END_METHOD


METHOD PRIVATE ShutdownMethodAccepted
VAR
    Accepted : BOOL;
END_VAR

TEST('ShutdownMethodAccepted');

ShutdownMethod.BusyCalls := 0;
Accepted := ShutdownMethod.Shutdown();
AssertTrue(Condition := Accepted, Message := 'Shutdown() returns TRUE');
AssertEquals_INT(Expected := 1, Actual := ShutdownMethod.Status.State, Message := 'REQUESTING before the block call');
ShutdownMethod();
AssertEquals_INT(Expected := 2, Actual := ShutdownMethod.Status.State, Message := 'SHUTTING_DOWN after the block call');
AssertEquals_INT(Expected := 1, Actual := ShutdownMethod.Requests, Message := 'one request sent');

TEST_FINISHED();
END_METHOD

END_FUNCTION_BLOCK

// ---- POUs/FB_PlcShutdownTestable.TcPOU

(*
    FB_PlcShutdown with a simulated operating system: SendRequest is
    overridden, so no shutdown request ever reaches the operating system.
    Used by FB_PlcShutdownTest and PRG_EXAMPLE.

    Simulation, like NT_Shutdown: a rising edge of Start sends a request.
    The request reports Busy for BusyCalls calls (counting the edge call),
    then completes, with an error if Fail is TRUE.
*)
FUNCTION_BLOCK FB_PlcShutdownTestable EXTENDS MBIDivB.FB_PlcShutdown
VAR_INPUT
    // Calls with Busy TRUE before the request completes.
    BusyCalls : INT := 2;
    // The request completes with ERR and FailErrorId.
    Fail : BOOL;
    FailErrorId : UDINT := 1793;
END_VAR
VAR_OUTPUT
    // Requests that would have reached the operating system.
    Requests : INT;
    // Delay of the last request, s.
    LastDelayS : UDINT;
END_VAR
VAR
    PreviousStart : BOOL;
    RemainingBusyCalls : INT;
END_VAR


SUPER^();


METHOD PROTECTED SendRequest
VAR_INPUT
    DelayS : UDINT;     // delay in seconds
    Start : BOOL;       // a rising edge sends the request
END_VAR
VAR_OUTPUT
    Busy : BOOL;        // request in progress
    Error : BOOL;       // request failed (valid when Busy is FALSE)
    ErrorId : UDINT;    // ADS error code of the failure
END_VAR

Busy := FALSE;
Error := FALSE;
ErrorId := 0;

IF Start AND NOT PreviousStart THEN
    Requests := Requests + 1;
    LastDelayS := DelayS;
    RemainingBusyCalls := BusyCalls;
END_IF
PreviousStart := Start;

IF NOT Start THEN
    RETURN;
END_IF
IF RemainingBusyCalls > 0 THEN
    RemainingBusyCalls := RemainingBusyCalls - 1;
    Busy := TRUE;
    RETURN;
END_IF
Error := Fail;
IF Fail THEN
    ErrorId := FailErrorId;
END_IF
END_METHOD

END_FUNCTION_BLOCK

// ---- Example/PRG_EXAMPLE.TcPOU

(*
    Example experiment program: every MBIDivB block, wired as an experiment's
    MAIN would do it. Driven over ADS from Linux by tools/ads_example.py
    (task 10.3 of openspec/changes/redesign-library-v1).

    No I/O is linked here. The program simulates the inputs instead:
    a sawtooth on Ai1, 1.0 V on Ai2 (the output of the amplifier Femto1),
    20 Hz flow sensor pulses, an EL2595 that reports "ready to activate",
    and valve switches that cycle through OPEN, BETWEEN, CLOSED, BETWEEN
    every 4000 cycles. Counter/timer channel 4 records the cycle number, so
    that the client can check the acquisition timing.

    Shutdown1 is FB_PlcShutdownTestable: its command handshake works, but no
    request ever reaches the operating system.

    Client-facing symbols: PRG_EXAMPLE.<instance>.Cmd/.Cfg/.Status, the data
    arrays PRG_EXAMPLE.Acq.Channel[c].Data and PRG_EXAMPLE.Ao1.Data, and
    PRG_EXAMPLE.StartAllTriggers for the group start of enabled triggers.
*)
PROGRAM PRG_EXAMPLE
VAR
    Ai1 : MBIDivB.FB_AnalogInput16;
    Ai2 : MBIDivB.FB_AnalogInput32;
    Acq : MBIDivB.FB_CounterTimer;
    Ao1 : MBIDivB.FB_AnalogOutput;
    Trig1 : MBIDivB.FB_MultiTrigger;
    Trig2 : MBIDivB.FB_MultiTrigger;
    Flow1 : MBIDivB.FB_FlowMeter;
    Shutter1 : MBIDivB.FB_ShutterControl;
    Led1 : MBIDivB.FB_LedControl;
    Femto1 : MBIDivB.FB_FemtoAmplifier;
    Valve1 : MBIDivB.FB_EndPositionSwitches;
    Shutdown1 : FB_PlcShutdownTestable;

    // Written TRUE by the client: starts all triggers with Cfg.Enabled.
    StartAllTriggers : BOOL;

    Initialized : BOOL;
    // Simulation: cycles since the PLC start.
    Cycle : UDINT;
END_VAR


// Initialization: terminal scaling
IF NOT Initialized THEN
    Initialized := TRUE;
    Ai1.SetScalePreset(Preset := MBIDivB.E_AiScalePreset.EL31XX_LEGACY, NominalFullScale := 10.0);
    Ai2.SetScalePreset(Preset := MBIDivB.E_AiScalePreset.ELM3XXX_EXTENDED, NominalFullScale := 10.0);
END_IF

// Simulated inputs (unlinked in this project)
Cycle := Cycle + 1;
Ai1.Raw := UDINT_TO_INT(Cycle MOD 1000) * 32;
Flow1.SensorInput := Cycle MOD 50 = 0;
Led1.StatusWord := 16#0001;
Ai2.Raw := 781250;  // 1.0 V with ELM3XXX_EXTENDED, 10 V
Valve1.OpenSwitch := Cycle MOD 4000 < 1500;
Valve1.ClosedSwitch := Cycle MOD 4000 >= 2000 AND Cycle MOD 4000 < 3500;

// Group start of the enabled triggers, before the trigger calls
IF StartAllTriggers THEN
    StartAllTriggers := FALSE;
    Trig1.StartIfEnabled();
    Trig2.StartIfEnabled();
END_IF

// Blocks
Ai1();
Ai2();
Femto1(Input := Ai2);   // after its input block
Ao1();
Trig1();
Trig2();
Flow1();
Shutter1();
Led1();
Valve1();
Shutdown1();

// Acquisition: channel inputs, then the block call, gated by trigger 1
Acq.Channel[1].Input := Ai1.Status.Value;
Acq.Channel[2].Input := Ao1.Status.Value;
Acq.Channel[3].Input := Flow1.Status.FlowRate;
Acq.Channel[4].Input := UDINT_TO_REAL(Cycle);
Acq(Gate := Trig1.Status.Output);

END_PROGRAM
